	IF pSpan <> 0 THEN
		THIS^.AssertEquals_UDINT(2, pSpan^.links.count, 'Expected two links');
		THIS^.AssertTrue(pSpan^.parentSpanId = 0, 'Expected a link not to make the span a child');
		pSpan^.links.reset();
		pLink := pSpan^.links.next();
		THIS^.AssertTrue(
			pLink <> 0 AND_THEN pTrigger <> 0 AND_THEN MEMCMP(ADR(pLink^.spanId^.bytes), ADR(pTrigger^.spanId^.bytes), SIZEOF(spanId.bytes)) = 0,
			'Expected the first link to point at the trigger span'
		);
		pLink := pSpan^.links.next();
		THIS^.AssertTrue(pLink <> 0 AND_THEN pLink^.traceId^.bytes[0] = 16#AA, 'Expected the second link to point at the remote trace');
		pSpan^.delete(pSelf:=pSpan);
	END_IF
	IF pTrigger <> 0 THEN pTrigger^.delete(pSelf:=pTrigger); END_IF
TcUnit.TEST_FINISHED();
END_METHOD

(* A null or all zero link context fails the chain, and build then releases the span. *)
METHOD testRejectsInvalidLink : REFERENCE TO FB_Test
VAR
	resource: FB_Resource('');
	idGenerator: FB_MockIdGenerator;
	provider: FB_TracerProvider(resource:=resource, idGenerator:=idGenerator, sampler:=TcOtlp_GVL.defaultSampler);
	scope: FB_InstrumentationScope('tracer.test', '1.0.0', '');
	tracer: FB_Tracer(scope:=scope, provider:=provider);
	pSpan: POINTER TO FB_Span;
	pZero: POINTER TO FB_SpanContext;
	traceId: FB_TraceId;
	spanId: FB_SpanId;
	success: BOOL;
	reason: E_TracerFailureReason;
END_VAR
TcUnit.TEST('testRejectsInvalidLink');
	success := tracer.startSpan(name:='work').addLink(pContext:=0).build(pDest:=pSpan, failureReason=>reason);
	THIS^.AssertFalse(success, 'Expected a null link context to fail the chain');
	THIS^.AssertEquals_UDINT(TO_UDINT(E_TracerFailureReason.LINK_CONTEXT_POINTER_NULL), TO_UDINT(reason), 'Expected LINK_CONTEXT_POINTER_NULL');
	THIS^.AssertTrue(pSpan = 0, 'Expected no span');

	ContextFactory.buildContext(pDest:=pZero, pTraceId:=ADR(traceId), pSpanId:=ADR(spanId), pTraceState:=0, traceFlags:=0);
	success := tracer.startSpan(name:='work').addLink(pContext:=pZero).build(pDest:=pSpan, failureReason=>reason);
	THIS^.AssertFalse(success, 'Expected an all zero link context to fail the chain');
	THIS^.AssertEquals_UDINT(TO_UDINT(E_TracerFailureReason.LINK_CONTEXT_INVALID), TO_UDINT(reason), 'Expected LINK_CONTEXT_INVALID');
	THIS^.AssertTrue(pSpan = 0, 'Expected no span');

	IF pZero <> 0 THEN pZero^.delete(pSelf:=pZero); END_IF
	IF pSpan <> 0 THEN pSpan^.delete(pSelf:=pSpan); END_IF
TcUnit.TEST_FINISHED();
END_METHOD

END_FUNCTION_BLOCK

// ---- TEST/TRACING/PROCESSOR/FB_SpanProcessor_ForInspection.TcPOU
(* Processor test double that counts what the simple processor does with each span. *)
FUNCTION_BLOCK FB_SpanProcessor_ForInspection EXTENDS FB_SpanProcessor_Simple
VAR_OUTPUT
	enrichedCount: UDINT;
	exportedCount: UDINT;
	tickCount: UDINT;
	enrichedBeforeExport: BOOL;
	lastSpanName: T_MaxString;
END_VAR

METHOD enrich
VAR_IN_OUT
	span: FB_Span;
END_VAR
THIS^.enrichedCount := THIS^.enrichedCount + 1;
END_METHOD

METHOD export
VAR_INPUT
	span: REFERENCE TO FB_Span;
END_VAR
THIS^.exportedCount := THIS^.exportedCount + 1;
THIS^.enrichedBeforeExport := THIS^.enrichedCount = THIS^.exportedCount;
IF span.name <> 0 AND_THEN span.name^.pString <> 0 THEN
	THIS^.lastSpanName := span.name^.pString^;
END_IF
END_METHOD

METHOD tick
THIS^.tickCount := THIS^.tickCount + 1;
END_METHOD

END_FUNCTION_BLOCK

// ---- TEST/TRACING/SPAN/FB_TestSpanQueue.TcPOU
(* Tests FB_SpanQueue ordering, its bound, and the ownership hand-off on push and pop.

   The spans are opaque queue nodes: the queue only moves and releases pointers, so the tests
   allocate bare spans with __NEW instead of building them through FB_Tracer. *)
FUNCTION_BLOCK FB_TestSpanQueue EXTENDS FB_TestSuite

THIS^.testPushPopIsFifo();
THIS^.testPushDropsOldestWhenFull();
THIS^.testPopIntoAssignedDestinationFails();
THIS^.testCursorWalksWithoutTakingOwnership();
THIS^.testTransferToMovesOldestSpans();
THIS^.testTransferToRejectsInvalidDestination();
THIS^.testRotateMovesOldestToBack();

(* push takes ownership and clears the caller's pointer; pop returns spans oldest first. *)
METHOD testPushPopIsFifo : REFERENCE TO FB_Test
VAR
	queue: FB_SpanQueue(maxCount:=4);
	pFirst: POINTER TO FB_Span;
	pSecond: POINTER TO FB_Span;
	pExpectedFirst: POINTER TO FB_Span;
	pExpectedSecond: POINTER TO FB_Span;
	pPopped: POINTER TO FB_Span;
	reason: E_SpanQueueFailureReason;
END_VAR
TcUnit.TEST('testPushPopIsFifo');
	pFirst := __NEW(FB_Span);  // opaque queue node: the queue needs no span identity
	pSecond := __NEW(FB_Span);
	pExpectedFirst := pFirst;
	pExpectedSecond := pSecond;

	THIS^.AssertTrue(queue.push(pValue:=pFirst, failureReason=>reason), 'Expected the first push to succeed');
	THIS^.AssertTrue(queue.push(pValue:=pSecond, failureReason=>reason), 'Expected the second push to succeed');
	THIS^.AssertTrue(pFirst = 0 AND pSecond = 0, 'Expected push to clear the caller$'s pointers');
	THIS^.AssertEquals_UDINT(2, queue.count, 'Expected two queued spans');

	THIS^.AssertTrue(queue.pop(pValue:=pPopped, failureReason=>reason), 'Expected the first pop to succeed');
	THIS^.AssertTrue(pPopped = pExpectedFirst, 'Expected the oldest span first');
	IF pPopped <> 0 THEN pPopped^.delete(pSelf:=pPopped); END_IF

	THIS^.AssertTrue(queue.pop(pValue:=pPopped, failureReason=>reason), 'Expected the second pop to succeed');
	THIS^.AssertTrue(pPopped = pExpectedSecond, 'Expected the newer span second');
	IF pPopped <> 0 THEN pPopped^.delete(pSelf:=pPopped); END_IF

	THIS^.AssertFalse(queue.pop(pValue:=pPopped, failureReason=>reason), 'Expected pop on an empty queue to fail');
	THIS^.AssertEquals_UDINT(
		TO_UDINT(E_SpanQueueFailureReason.QUEUE_EMPTY),
		TO_UDINT(reason),
		'Expected QUEUE_EMPTY'
	);
	THIS^.AssertEquals_UDINT(0, queue.count, 'Expected the queue to be empty');
TcUnit.TEST_FINISHED();
END_METHOD

(* A full queue releases its oldest span to make room and counts the drop. *)
METHOD testPushDropsOldestWhenFull : REFERENCE TO FB_Test
VAR
	queue: FB_SpanQueue(maxCount:=1);
	pOld: POINTER TO FB_Span;
	pNew: POINTER TO FB_Span;
	pExpected: POINTER TO FB_Span;
	pPopped: POINTER TO FB_Span;
	reason: E_SpanQueueFailureReason;
END_VAR
TcUnit.TEST('testPushDropsOldestWhenFull');
	pOld := __NEW(FB_Span);  // opaque queue node: the queue needs no span identity
	pNew := __NEW(FB_Span);
	pExpected := pNew;

	queue.push(pValue:=pOld, failureReason=>reason);
	THIS^.AssertTrue(queue.push(pValue:=pNew, failureReason=>reason), 'Expected push to a full queue to succeed');
	THIS^.AssertEquals_UDINT(1, queue.count, 'Expected the bound to hold');
	THIS^.AssertEquals_UDINT(1, queue.droppedCount, 'Expected one dropped span');

	queue.pop(pValue:=pPopped, failureReason=>reason);
	THIS^.AssertTrue(pPopped = pExpected, 'Expected the newest span to be kept');
	IF pPopped <> 0 THEN pPopped^.delete(pSelf:=pPopped); END_IF
TcUnit.TEST_FINISHED();
END_METHOD

(* pop never overwrites a pointer the caller already owns, and free releases what is left. *)
METHOD testPopIntoAssignedDestinationFails : REFERENCE TO FB_Test
VAR
	queue: FB_SpanQueue(maxCount:=4);
	pQueued: POINTER TO FB_Span;
	pOwned: POINTER TO FB_Span;
	pExpected: POINTER TO FB_Span;
	reason: E_SpanQueueFailureReason;
END_VAR
TcUnit.TEST('testPopIntoAssignedDestinationFails');
	pQueued := __NEW(FB_Span);  // opaque queue node: the queue needs no span identity
	pOwned := __NEW(FB_Span);  // held by the caller, so pop must not overwrite it
	pExpected := pOwned;
	queue.push(pValue:=pQueued, failureReason=>reason);

	THIS^.AssertFalse(queue.pop(pValue:=pOwned, failureReason=>reason), 'Expected pop into an assigned pointer to fail');
	THIS^.AssertEquals_UDINT(
		TO_UDINT(E_SpanQueueFailureReason.DESTINATION_ALREADY_ASSIGNED),
		TO_UDINT(reason),
		'Expected DESTINATION_ALREADY_ASSIGNED'
	);
	THIS^.AssertTrue(pOwned = pExpected, 'Expected the destination to be left alone');
	THIS^.AssertEquals_UDINT(1, queue.count, 'Expected the span to stay queued');

	THIS^.AssertTrue(queue.free(), 'Expected free to release every span');
	THIS^.AssertEquals_UDINT(0, queue.count, 'Expected an empty queue after free');
	IF pOwned <> 0 THEN pOwned^.delete(pSelf:=pOwned); END_IF
TcUnit.TEST_FINISHED();
END_METHOD

(* reset and next walk the spans oldest first and leave them queued; pop keeps the cursor valid. *)
METHOD testCursorWalksWithoutTakingOwnership : REFERENCE TO FB_Test
VAR
	queue: FB_SpanQueue(maxCount:=4);
	pFirst: POINTER TO FB_Span;
	pSecond: POINTER TO FB_Span;
	pExpectedFirst: POINTER TO FB_Span;
	pExpectedSecond: POINTER TO FB_Span;
	pPopped: POINTER TO FB_Span;
END_VAR
TcUnit.TEST('testCursorWalksWithoutTakingOwnership');
	pFirst := __NEW(FB_Span);  // opaque queue node: the queue needs no span identity
	pSecond := __NEW(FB_Span);
	pExpectedFirst := pFirst;
	pExpectedSecond := pSecond;
	queue.push(pValue:=pFirst);
	queue.push(pValue:=pSecond);

	queue.reset();
	THIS^.AssertTrue(queue.next() = pExpectedFirst, 'Expected the oldest span first');
	THIS^.AssertTrue(queue.next() = pExpectedSecond, 'Expected the second span next');
	THIS^.AssertTrue(queue.next() = 0, 'Expected 0 after the last span');
	THIS^.AssertEquals_UDINT(2, queue.count, 'Expected the walk to leave both spans queued');

	// popping the node under the cursor moves the cursor to the new head
	queue.reset();
	queue.pop(pValue:=pPopped);
	THIS^.AssertTrue(queue.next() = pExpectedSecond, 'Expected the cursor to move past the popped span');

	IF pPopped <> 0 THEN pPopped^.delete(pSelf:=pPopped); END_IF
	queue.free();
	queue.reset();
	THIS^.AssertTrue(queue.next() = 0, 'Expected an empty walk after free');
TcUnit.TEST_FINISHED();
END_METHOD

(* transferTo moves the oldest spans, up to the destination's bound, without copying them. *)
METHOD testTransferToMovesOldestSpans : REFERENCE TO FB_Test
VAR
	source: FB_SpanQueue(maxCount:=4);
	destination: FB_SpanQueue(maxCount:=2);
	p: POINTER TO FB_Span;
	pFirst: POINTER TO FB_Span;
	pSecond: POINTER TO FB_Span;
	pThird: POINTER TO FB_Span;
	pPopped: POINTER TO FB_Span;
	reason: E_SpanQueueFailureReason;
END_VAR
TcUnit.TEST('testTransferToMovesOldestSpans');
	// opaque queue nodes: the queue needs no span identity
	p := __NEW(FB_Span); pFirst := p; source.push(pValue:=p, failureReason=>reason);
	p := __NEW(FB_Span); pSecond := p; source.push(pValue:=p, failureReason=>reason);
	p := __NEW(FB_Span); pThird := p; source.push(pValue:=p, failureReason=>reason);

	// ask for more than the destination's bound of 2 and more than the source holds
	THIS^.AssertTrue(source.transferTo(destination:=destination, count:=5, failureReason=>reason), 'Expected transferTo to succeed');
	THIS^.AssertEquals_UDINT(2, destination.count, 'Expected the destination bound to hold');
	THIS^.AssertEquals_UDINT(1, source.count, 'Expected one span left behind');

	destination.pop(pValue:=pPopped, failureReason=>reason);
	THIS^.AssertTrue(pPopped = pFirst, 'Expected the oldest span first');
	IF pPopped <> 0 THEN pPopped^.delete(pSelf:=pPopped); END_IF
	destination.pop(pValue:=pPopped, failureReason=>reason);
	THIS^.AssertTrue(pPopped = pSecond, 'Expected the second span next');
	IF pPopped <> 0 THEN pPopped^.delete(pSelf:=pPopped); END_IF
	source.pop(pValue:=pPopped, failureReason=>reason);
	THIS^.AssertTrue(pPopped = pThird, 'Expected the newest span to stay in the source');
	IF pPopped <> 0 THEN pPopped^.delete(pSelf:=pPopped); END_IF

	THIS^.AssertTrue(source.transferTo(destination:=destination, count:=1, failureReason=>reason), 'Expected an empty transfer to succeed');
	THIS^.AssertEquals_UDINT(0, destination.count, 'Expected nothing to move from an empty queue');
	source.free();
	destination.free();
TcUnit.TEST_FINISHED();
END_METHOD

(* transferTo refuses itself and a non-empty destination, and moves nothing. *)
METHOD testTransferToRejectsInvalidDestination : REFERENCE TO FB_Test
VAR
	source: FB_SpanQueue(maxCount:=4);
	destination: FB_SpanQueue(maxCount:=4);
	p: POINTER TO FB_Span;
	reason: E_SpanQueueFailureReason;
END_VAR
TcUnit.TEST('testTransferToRejectsInvalidDestination');
	// opaque queue nodes: the queue needs no span identity
	p := __NEW(FB_Span); source.push(pValue:=p, failureReason=>reason);
	p := __NEW(FB_Span); destination.push(pValue:=p, failureReason=>reason);  // makes the destination non-empty

	THIS^.AssertFalse(source.transferTo(destination:=source, count:=1, failureReason=>reason), 'Expected a self transfer to fail');
	THIS^.AssertEquals_UDINT(
		TO_UDINT(E_SpanQueueFailureReason.SELF_TRANSFER_NOT_ALLOWED),
		TO_UDINT(reason),
		'Expected SELF_TRANSFER_NOT_ALLOWED'
	);
	THIS^.AssertFalse(source.transferTo(destination:=destination, count:=1, failureReason=>reason), 'Expected a non-empty destination to fail');
	THIS^.AssertEquals_UDINT(
		TO_UDINT(E_SpanQueueFailureReason.DESTINATION_NOT_EMPTY),
		TO_UDINT(reason),
		'Expected DESTINATION_NOT_EMPTY'
	);
	THIS^.AssertTrue(source.count = 1 AND destination.count = 1, 'Expected both queues to be unchanged');
	source.free();
	destination.free();
TcUnit.TEST_FINISHED();
END_METHOD

(* rotate moves the oldest span to the back without releasing it, and fails on an empty queue. *)
METHOD testRotateMovesOldestToBack : REFERENCE TO FB_Test
VAR
	queue: FB_SpanQueue(maxCount:=0);  // 0 means the default bound, MAX_LOOP_COUNT
	pSpan: POINTER TO FB_Span;
	pFirst: POINTER TO FB_Span;
	pSecond: POINTER TO FB_Span;
	pPopped: POINTER TO FB_Span;
	reason: E_SpanQueueFailureReason;
END_VAR
TcUnit.TEST('testRotateMovesOldestToBack');
	THIS^.AssertFalse(queue.rotate(failureReason=>reason), 'Expected rotate on an empty queue to fail');
	THIS^.AssertEquals_UDINT(TO_UDINT(E_SpanQueueFailureReason.QUEUE_EMPTY), TO_UDINT(reason), 'Expected QUEUE_EMPTY');

	pSpan := __NEW(FB_Span);  // opaque queue node: the queue needs no span identity
	pFirst := pSpan;
	queue.push(pValue:=pSpan);
	pSpan := __NEW(FB_Span);
	pSecond := pSpan;
	queue.push(pValue:=pSpan);

	THIS^.AssertTrue(queue.rotate(failureReason=>reason), 'Expected rotate to succeed');
	THIS^.AssertEquals_UDINT(2, queue.count, 'Expected rotate to keep both spans');
	THIS^.AssertTrue(queue.next() = pSecond, 'Expected the cursor at the new head');
	queue.pop(pValue:=pPopped);
	THIS^.AssertTrue(pPopped = pSecond, 'Expected the second span first after a rotate');
	IF pPopped <> 0 THEN pPopped^.delete(pSelf:=pPopped); END_IF
	queue.pop(pValue:=pPopped);
	THIS^.AssertTrue(pPopped = pFirst, 'Expected the rotated span last');
	IF pPopped <> 0 THEN pPopped^.delete(pSelf:=pPopped); END_IF
	queue.free();
TcUnit.TEST_FINISHED();
END_METHOD

END_FUNCTION_BLOCK

// ---- TEST/TRACING/PROCESSOR/FB_TestSpanProcessors.TcPOU
(* Tests FB_SpanProcessor_Simple and FB_SpanProcessor_Batch and their hand-off to an exporter. *)
FUNCTION_BLOCK FB_TestSpanProcessors EXTENDS FB_TestSuite
VAR
	// kept across scans by testBatchExportsAfterScheduledDelay
	_resource: FB_Resource('');
	_idGenerator: FB_MockIdGenerator;
	_provider: FB_TracerProvider_ForInspection(resource:=_resource, idGenerator:=_idGenerator, sampler:=TcOtlp_GVL.defaultSampler);
	_scope: FB_InstrumentationScope('tracer.test', '1.0.0', '');
	_tracer: FB_Tracer(scope:=_scope, provider:=_provider);
	_exporter: FB_SpanExporter_ForInspection;
	_processor: FB_SpanProcessor_Batch(maxQueueSize:=10, scheduledDelayMillis:=50, maxExportBatchSize:=10, exporter:=_exporter);
END_VAR

THIS^.testSimpleEnrichesThenExports();
THIS^.testSimpleHandsCloneToExporter();
THIS^.testSimpleDropsSpanWhenExporterBusy();
THIS^.testBatchWaitsForFullBatch();
THIS^.testBatchKeepsSpansWhileExporterBusy();
THIS^.testBatchDropsOldestWhenFull();
THIS^.testBatchIgnoresSpansWithoutExporter();
THIS^.testBatchExportsAfterScheduledDelay();

(* The simple processor enriches each span and then exports it, once per span. *)
METHOD testSimpleEnrichesThenExports : REFERENCE TO FB_Test
VAR
	resource: FB_Resource('');
	idGenerator: FB_MockIdGenerator;
	provider: FB_TracerProvider_ForInspection(resource:=resource, idGenerator:=idGenerator, sampler:=TcOtlp_GVL.defaultSampler);
	scope: FB_InstrumentationScope('tracer.test', '1.0.0', '');
	tracer: FB_Tracer(scope:=scope, provider:=provider);
	processor: FB_SpanProcessor_ForInspection(exporter:=0);
	pSpan: POINTER TO FB_Span;
END_VAR
TcUnit.TEST('testSimpleEnrichesThenExports');
	tracer.startSpan(name:='work').build(pDest:=pSpan);
	THIS^.AssertTrue(pSpan <> 0, 'Expected the span to build');
	IF pSpan <> 0 THEN
		processor.onEnd(pSpan^);
		pSpan^.delete(pSelf:=pSpan);
	END_IF
	THIS^.AssertEquals_UDINT(1, processor.enrichedCount, 'Expected one enrich');
	THIS^.AssertEquals_UDINT(1, processor.exportedCount, 'Expected one export');
	THIS^.AssertTrue(processor.enrichedBeforeExport, 'Expected enrich to run before export');
	THIS^.AssertEquals_STRING('work', processor.lastSpanName, 'Expected the span to be exported');
TcUnit.TEST_FINISHED();
END_METHOD

(* The simple processor gives the exporter a clone, which outlives the span the provider releases. *)
METHOD testSimpleHandsCloneToExporter : REFERENCE TO FB_Test
VAR
	resource: FB_Resource('');
	idGenerator: FB_MockIdGenerator;
	provider: FB_TracerProvider_ForInspection(resource:=resource, idGenerator:=idGenerator, sampler:=TcOtlp_GVL.defaultSampler);
	scope: FB_InstrumentationScope('tracer.test', '1.0.0', '');
	tracer: FB_Tracer(scope:=scope, provider:=provider);
	exporter: FB_SpanExporter_ForInspection;
	processor: FB_SpanProcessor_Simple(exporter:=exporter);
	pSpan: POINTER TO FB_Span;
	pSource: POINTER TO FB_Span;
	pHeld: POINTER TO FB_Span;
END_VAR
TcUnit.TEST('testSimpleHandsCloneToExporter');
	tracer.startSpan(name:='work').build(pDest:=pSpan);
	THIS^.AssertTrue(pSpan <> 0, 'Expected the span to build');
	IF pSpan <> 0 THEN
		pSource := pSpan;
		processor.onEnd(pSpan^);
		pSpan^.delete(pSelf:=pSpan);
	END_IF
	THIS^.AssertEquals_UDINT(1, exporter.exportCount, 'Expected one export');
	THIS^.AssertEquals_UDINT(1, exporter.lastBatchCount, 'Expected a batch of one');
	pHeld := exporter.heldSpan();
	THIS^.AssertTrue(pHeld <> 0 AND_THEN pHeld <> pSource, 'Expected the exporter to hold a clone');
	IF pHeld <> 0 AND_THEN pHeld^.name <> 0 THEN
		THIS^.AssertEquals_STRING('work', pHeld^.name^.pString^, 'Expected the clone to outlive the source');
	END_IF
	processor.tick();
	THIS^.AssertEquals_UDINT(1, exporter.tickCount, 'Expected tick to reach the exporter');
	exporter.free();
TcUnit.TEST_FINISHED();
END_METHOD

(* A busy exporter is not offered the span, and nothing is kept for later. *)
METHOD testSimpleDropsSpanWhenExporterBusy : REFERENCE TO FB_Test
VAR
	resource: FB_Resource('');
	idGenerator: FB_MockIdGenerator;
	provider: FB_TracerProvider_ForInspection(resource:=resource, idGenerator:=idGenerator, sampler:=TcOtlp_GVL.defaultSampler);
	scope: FB_InstrumentationScope('tracer.test', '1.0.0', '');
	tracer: FB_Tracer(scope:=scope, provider:=provider);
	exporter: FB_SpanExporter_ForInspection;
	processor: FB_SpanProcessor_Simple(exporter:=exporter);
	pSpan: POINTER TO FB_Span;
END_VAR
TcUnit.TEST('testSimpleDropsSpanWhenExporterBusy');
	exporter.busy := TRUE;
	tracer.startSpan(name:='work').build(pDest:=pSpan);
	IF pSpan <> 0 THEN
		processor.onEnd(pSpan^);
		pSpan^.delete(pSelf:=pSpan);
	END_IF
	THIS^.AssertEquals_UDINT(0, exporter.exportCount, 'Expected no export while busy');
	THIS^.AssertEquals_UDINT(0, exporter.callsWhileBusy, 'Expected the processor not to call a busy exporter');
	THIS^.AssertTrue(exporter.heldSpan() = 0, 'Expected the exporter to hold nothing');
TcUnit.TEST_FINISHED();
END_METHOD

(* Ended spans are only queued; a full batch goes out on the next tick without waiting for the delay. *)
METHOD testBatchWaitsForFullBatch : REFERENCE TO FB_Test
VAR
	resource: FB_Resource('');
	idGenerator: FB_MockIdGenerator;
	provider: FB_TracerProvider_ForInspection(resource:=resource, idGenerator:=idGenerator, sampler:=TcOtlp_GVL.defaultSampler);
	scope: FB_InstrumentationScope('tracer.test', '1.0.0', '');
	tracer: FB_Tracer(scope:=scope, provider:=provider);
	exporter: FB_SpanExporter_ForInspection;
	processor: FB_SpanProcessor_Batch(maxQueueSize:=10, scheduledDelayMillis:=60000, maxExportBatchSize:=3, exporter:=exporter);
	pSpan: POINTER TO FB_Span;
END_VAR
TcUnit.TEST('testBatchWaitsForFullBatch');
	tracer.startSpan(name:='a').build(pDest:=pSpan);
	IF pSpan <> 0 THEN
		processor.onEnd(pSpan^);
		pSpan^.delete(pSelf:=pSpan);
	END_IF
	tracer.startSpan(name:='b').build(pDest:=pSpan);
	IF pSpan <> 0 THEN
		processor.onEnd(pSpan^);
		pSpan^.delete(pSelf:=pSpan);
	END_IF
	THIS^.AssertEquals_UDINT(0, exporter.exportCount, 'Expected onEnd not to export');
	THIS^.AssertEquals_UDINT(2, processor.queuedCount, 'Expected two queued spans');
	processor.tick();
	THIS^.AssertEquals_UDINT(0, exporter.exportCount, 'Expected no export before a full batch or the delay');
	THIS^.AssertEquals_UDINT(1, exporter.tickCount, 'Expected tick to reach the exporter');
	tracer.startSpan(name:='c').build(pDest:=pSpan);
	IF pSpan <> 0 THEN
		processor.onEnd(pSpan^);
		pSpan^.delete(pSelf:=pSpan);
	END_IF
	processor.tick();
	THIS^.AssertEquals_UDINT(1, exporter.exportCount, 'Expected one export for the full batch');
	THIS^.AssertEquals_UDINT(3, exporter.lastBatchCount, 'Expected the three spans in one batch');
	THIS^.AssertEquals_UDINT(0, processor.queuedCount, 'Expected the queue to be empty');
	THIS^.AssertEquals_UDINT(0, processor.droppedCount, 'Expected nothing dropped');
	exporter.free();
	processor.free();
TcUnit.TEST_FINISHED();
END_METHOD

(* Spans that end while the exporter is busy stay queued and are exported once it is idle. *)
METHOD testBatchKeepsSpansWhileExporterBusy : REFERENCE TO FB_Test
VAR
	resource: FB_Resource('');
	idGenerator: FB_MockIdGenerator;
	provider: FB_TracerProvider_ForInspection(resource:=resource, idGenerator:=idGenerator, sampler:=TcOtlp_GVL.defaultSampler);
	scope: FB_InstrumentationScope('tracer.test', '1.0.0', '');
	tracer: FB_Tracer(scope:=scope, provider:=provider);
	exporter: FB_SpanExporter_ForInspection;
	processor: FB_SpanProcessor_Batch(maxQueueSize:=10, scheduledDelayMillis:=60000, maxExportBatchSize:=1, exporter:=exporter);
	pSpan: POINTER TO FB_Span;
	pHeld: POINTER TO FB_Span;
END_VAR
TcUnit.TEST('testBatchKeepsSpansWhileExporterBusy');
	exporter.busy := TRUE;
	tracer.startSpan(name:='first').build(pDest:=pSpan);
	IF pSpan <> 0 THEN
		processor.onEnd(pSpan^);
		pSpan^.delete(pSelf:=pSpan);
	END_IF
	tracer.startSpan(name:='second').build(pDest:=pSpan);
	IF pSpan <> 0 THEN
		processor.onEnd(pSpan^);
		pSpan^.delete(pSelf:=pSpan);
	END_IF
	processor.tick();
	THIS^.AssertEquals_UDINT(0, exporter.exportCount, 'Expected no export while busy');
	THIS^.AssertEquals_UDINT(0, exporter.callsWhileBusy, 'Expected the processor not to call a busy exporter');
	THIS^.AssertEquals_UDINT(2, processor.queuedCount, 'Expected both spans kept');

	exporter.busy := FALSE;
	processor.tick();
	THIS^.AssertEquals_UDINT(1, exporter.exportCount, 'Expected an export once idle');
	THIS^.AssertEquals_UDINT(1, exporter.lastBatchCount, 'Expected a batch of maxExportBatchSize');
	pHeld := exporter.heldSpan();
	IF pHeld <> 0 AND_THEN pHeld^.name <> 0 THEN
		THIS^.AssertEquals_STRING('first', pHeld^.name^.pString^, 'Expected the oldest span first');
	ELSE
		THIS^.AssertTrue(FALSE, 'Expected the exporter to hold a span');
	END_IF
	THIS^.AssertEquals_UDINT(1, processor.queuedCount, 'Expected the newer span to wait');

	processor.tick();
	THIS^.AssertEquals_UDINT(2, exporter.exportCount, 'Expected the second span on the next tick');
	pHeld := exporter.heldSpan();
	IF pHeld <> 0 AND_THEN pHeld^.name <> 0 THEN
		THIS^.AssertEquals_STRING('second', pHeld^.name^.pString^, 'Expected the newer span second');
	END_IF
	THIS^.AssertEquals_UDINT(0, processor.droppedCount, 'Expected nothing dropped');
	exporter.free();
	processor.free();
TcUnit.TEST_FINISHED();
END_METHOD

(* A full queue drops its oldest span for the newest and counts it. *)
METHOD testBatchDropsOldestWhenFull : REFERENCE TO FB_Test
VAR
	resource: FB_Resource('');
	idGenerator: FB_MockIdGenerator;
	provider: FB_TracerProvider_ForInspection(resource:=resource, idGenerator:=idGenerator, sampler:=TcOtlp_GVL.defaultSampler);
	scope: FB_InstrumentationScope('tracer.test', '1.0.0', '');
	tracer: FB_Tracer(scope:=scope, provider:=provider);
	exporter: FB_SpanExporter_ForInspection;
	processor: FB_SpanProcessor_Batch(maxQueueSize:=2, scheduledDelayMillis:=60000, maxExportBatchSize:=2, exporter:=exporter);
	pSpan: POINTER TO FB_Span;
	pHeld: POINTER TO FB_Span;
END_VAR
TcUnit.TEST('testBatchDropsOldestWhenFull');
	exporter.busy := TRUE;
	tracer.startSpan(name:='a').build(pDest:=pSpan);
	IF pSpan <> 0 THEN
		processor.onEnd(pSpan^);
		pSpan^.delete(pSelf:=pSpan);
	END_IF
	tracer.startSpan(name:='b').build(pDest:=pSpan);
	IF pSpan <> 0 THEN
		processor.onEnd(pSpan^);
		pSpan^.delete(pSelf:=pSpan);
	END_IF
	tracer.startSpan(name:='c').build(pDest:=pSpan);
	IF pSpan <> 0 THEN
		processor.onEnd(pSpan^);
		pSpan^.delete(pSelf:=pSpan);
	END_IF
	THIS^.AssertEquals_UDINT(2, processor.queuedCount, 'Expected the queue to stay at maxQueueSize');
	THIS^.AssertEquals_UDINT(1, processor.droppedCount, 'Expected one dropped span');
	processor.tick();
	THIS^.AssertEquals_UDINT(0, exporter.callsWhileBusy, 'Expected the processor not to call a busy exporter with a full batch');
	exporter.busy := FALSE;
	processor.tick();
	THIS^.AssertEquals_UDINT(2, exporter.lastBatchCount, 'Expected the two kept spans');
	pHeld := exporter.heldSpan();
	IF pHeld <> 0 AND_THEN pHeld^.name <> 0 THEN
		THIS^.AssertEquals_STRING('b', pHeld^.name^.pString^, 'Expected the oldest span to be the one dropped');
	ELSE
		THIS^.AssertTrue(FALSE, 'Expected the exporter to hold a span');
	END_IF
	exporter.free();
	processor.free();
TcUnit.TEST_FINISHED();
END_METHOD

(* With no exporter the processor keeps nothing. *)
METHOD testBatchIgnoresSpansWithoutExporter : REFERENCE TO FB_Test
VAR
	resource: FB_Resource('');
	idGenerator: FB_MockIdGenerator;
	provider: FB_TracerProvider_ForInspection(resource:=resource, idGenerator:=idGenerator, sampler:=TcOtlp_GVL.defaultSampler);
	scope: FB_InstrumentationScope('tracer.test', '1.0.0', '');
	tracer: FB_Tracer(scope:=scope, provider:=provider);
	exporter: FB_SpanExporter_ForInspection;
	processor: FB_SpanProcessor_Batch(maxQueueSize:=10, scheduledDelayMillis:=0, maxExportBatchSize:=1, exporter:=0);
	pSpan: POINTER TO FB_Span;
END_VAR
TcUnit.TEST('testBatchIgnoresSpansWithoutExporter');
	tracer.startSpan(name:='work').build(pDest:=pSpan);
	IF pSpan <> 0 THEN
		processor.onEnd(pSpan^);
		pSpan^.delete(pSelf:=pSpan);
	END_IF
	processor.tick();
	THIS^.AssertEquals_UDINT(0, processor.queuedCount, 'Expected nothing queued');
TcUnit.TEST_FINISHED();
END_METHOD

(* A partial batch is exported once scheduledDelayMillis has passed, and not before. *)
METHOD testBatchExportsAfterScheduledDelay : REFERENCE TO FB_Test
VAR CONSTANT
	DELAY_MILLIS: UDINT := 50;  // matches _processor's scheduledDelayMillis
	MAX_CYCLES: UDINT := 1000;
END_VAR
VAR_INST
	_started: BOOL;
	_finished: BOOL;
	_cycles: UDINT;
	_startTime: ULINT;
END_VAR
VAR
	pSpan: POINTER TO FB_Span;
	elapsedMillis: ULINT;
END_VAR
TcUnit.TEST('testBatchExportsAfterScheduledDelay');
	IF _finished THEN
		RETURN;
	END_IF
	IF NOT _started THEN
		_tracer.startSpan(name:='work').build(pDest:=pSpan);
		IF pSpan <> 0 THEN
			_processor.onEnd(pSpan^);
			pSpan^.delete(pSelf:=pSpan);
		END_IF
		_startTime := F_GetSystemTime();
		_started := TRUE;
	END_IF

	_processor.tick();
	_cycles := _cycles + 1;
	IF _exporter.exportCount > 0 OR _cycles > MAX_CYCLES THEN
		elapsedMillis := (F_GetSystemTime() - _startTime) / 10000;  // 100 ns ticks
		THIS^.AssertEquals_UDINT(1, _exporter.exportCount, 'Expected the partial batch to be exported');
		THIS^.AssertEquals_UDINT(1, _exporter.lastBatchCount, 'Expected a batch of one');
		THIS^.AssertTrue(elapsedMillis >= DELAY_MILLIS - 1, 'Expected the export to wait for the delay');
		_exporter.free();
		_processor.free();
		_finished := TRUE;
		TcUnit.TEST_FINISHED();
	END_IF
END_METHOD

END_FUNCTION_BLOCK

// ---- TEST/TRACING/EXPORTING/FB_SpanExporter_ForInspection.TcPOU
(*
	Span exporter test double. It keeps each accepted batch until the next one or free, and is
	busy while busy is set. callsWhileBusy counts export calls made while busy, which a processor
	must never make.
*)
FUNCTION_BLOCK FB_SpanExporter_ForInspection EXTENDS FB_SpanExporter_Base
VAR_INPUT
	busy: BOOL;
END_VAR
VAR_OUTPUT
	exportCount: UDINT;
	lastBatchCount: UDINT;
	tickCount: UDINT;
	callsWhileBusy: UDINT;
END_VAR

METHOD export : BOOL
VAR_IN_OUT
	spans: FB_SpanQueue;
END_VAR
VAR_INPUT
	count: UDINT;
END_VAR
VAR_OUTPUT
	failureReason: E_SpanExporterFailureReason;
END_VAR
IF THIS^.isBusy() THEN
	THIS^.callsWhileBusy := THIS^.callsWhileBusy + 1;
END_IF
export := SUPER^.export(spans:=spans, count:=count, failureReason=>failureReason);
IF export THEN
	THIS^.exportCount := THIS^.exportCount + 1;
	THIS^.lastBatchCount := THIS^._spans.count;
	// nothing is delivered, so the batch stays held until the next one or free
	THIS^._exportActive := FALSE;
END_IF
END_METHOD

(* The oldest span of the held batch, borrowed; 0 when nothing is held. *)
METHOD heldSpan : POINTER TO FB_Span
THIS^._spans.reset();
heldSpan := THIS^._spans.next();
END_METHOD

METHOD isBusy : BOOL
isBusy := THIS^.busy;
END_METHOD

METHOD tick : BOOL
VAR_OUTPUT
	failureReason: E_SpanExporterFailureReason;
END_VAR
THIS^.tickCount := THIS^.tickCount + 1;
failureReason := E_SpanExporterFailureReason.NA;
tick := TRUE;
END_METHOD

END_FUNCTION_BLOCK

// ---- TEST/TRACING/PROVIDER/FB_TestTracerProvider.TcPOU
(* Tests FB_TracerProvider processor staging and the hand-over of ended spans in tick. *)
FUNCTION_BLOCK FB_TestTracerProvider EXTENDS FB_TestSuite

THIS^.testTickHandsSpansToEachProcessor();
THIS^.testStageProcessorIgnoresDuplicates();
THIS^.testTickWithoutProcessorsSucceeds();
THIS^.testProcessorsMustBeStagedEachScan();

(* Every staged processor receives every ended span once; tick then releases the spans. *)
METHOD testTickHandsSpansToEachProcessor : REFERENCE TO FB_Test
VAR
	resource: FB_Resource('');
	idGenerator: FB_MockIdGenerator;
	provider: FB_TracerProvider_ForInspection(resource:=resource, idGenerator:=idGenerator, sampler:=TcOtlp_GVL.defaultSampler);
	scope: FB_InstrumentationScope('tracer.test', '1.0.0', '');
	tracer: FB_Tracer(scope:=scope, provider:=provider);
	processorA: FB_SpanProcessor_ForInspection(exporter:=0);
	processorB: FB_SpanProcessor_ForInspection(exporter:=0);
	pSpan: POINTER TO FB_Span;
	success: BOOL;
	reason: E_TracerProviderFailureReason;
END_VAR
TcUnit.TEST('testTickHandsSpansToEachProcessor');
	provider.stageProcessor(processorA).stageProcessor(processorB);
	tracer.startSpan(name:='first').build(pDest:=pSpan);
	tracer.endSpan(pSpan:=pSpan);
	tracer.startSpan(name:='second').build(pDest:=pSpan);
	tracer.endSpan(pSpan:=pSpan);

	success := provider.tick(failureReason=>reason);
	THIS^.AssertTrue(success, 'Expected tick to succeed');
	THIS^.AssertEquals_UDINT(
		TO_UDINT(E_TracerProviderFailureReason.NA),
		TO_UDINT(reason),
		'Expected no failure reason on success'
	);
	THIS^.AssertEquals_UDINT(2, processorA.exportedCount, 'Expected processor A to get both spans');
	THIS^.AssertEquals_UDINT(2, processorB.exportedCount, 'Expected processor B to get both spans');
	THIS^.AssertEquals_STRING('second', processorA.lastSpanName, 'Expected the spans in the order they ended');
	THIS^.AssertEquals_UDINT(1, processorA.tickCount, 'Expected each processor to be ticked once');
	THIS^.AssertEquals_UDINT(0, provider.spans.count, 'Expected the queue to be empty');
	THIS^.AssertEquals_UDINT(0, provider.stagedProcessorCount, 'Expected the staged list to be cleared');
TcUnit.TEST_FINISHED();
END_METHOD

(* Staging the same processor twice gives it each span once. *)
METHOD testStageProcessorIgnoresDuplicates : REFERENCE TO FB_Test
VAR
	resource: FB_Resource('');
	idGenerator: FB_MockIdGenerator;
	provider: FB_TracerProvider_ForInspection(resource:=resource, idGenerator:=idGenerator, sampler:=TcOtlp_GVL.defaultSampler);
	scope: FB_InstrumentationScope('tracer.test', '1.0.0', '');
	tracer: FB_Tracer(scope:=scope, provider:=provider);
	processor: FB_SpanProcessor_ForInspection(exporter:=0);
	pSpan: POINTER TO FB_Span;
END_VAR
TcUnit.TEST('testStageProcessorIgnoresDuplicates');
	provider.stageProcessor(processor).stageProcessor(processor);
	THIS^.AssertEquals_UDINT(1, provider.stagedProcessorCount, 'Expected the duplicate to be ignored');

	tracer.startSpan(name:='work').build(pDest:=pSpan);
	tracer.endSpan(pSpan:=pSpan);
	provider.tick();
	THIS^.AssertEquals_UDINT(1, processor.exportedCount, 'Expected the span exactly once');
TcUnit.TEST_FINISHED();
END_METHOD

(* With no processors staged, tick releases the queued spans and still succeeds. *)
METHOD testTickWithoutProcessorsSucceeds : REFERENCE TO FB_Test
VAR
	resource: FB_Resource('');
	idGenerator: FB_MockIdGenerator;
	provider: FB_TracerProvider_ForInspection(resource:=resource, idGenerator:=idGenerator, sampler:=TcOtlp_GVL.defaultSampler);
	scope: FB_InstrumentationScope('tracer.test', '1.0.0', '');
	tracer: FB_Tracer(scope:=scope, provider:=provider);
	pSpan: POINTER TO FB_Span;
	success: BOOL;
END_VAR
TcUnit.TEST('testTickWithoutProcessorsSucceeds');
	tracer.startSpan(name:='work').build(pDest:=pSpan);
	tracer.endSpan(pSpan:=pSpan);
	THIS^.AssertEquals_UDINT(1, provider.spans.count, 'Expected the span to be queued');

	success := provider.tick();
	THIS^.AssertTrue(success, 'Expected tick to succeed');
	THIS^.AssertEquals_UDINT(0, provider.spans.count, 'Expected tick to release the span');
TcUnit.TEST_FINISHED();
END_METHOD

(* tick clears the staged list, so a processor that is not staged again gets nothing. *)
METHOD testProcessorsMustBeStagedEachScan : REFERENCE TO FB_Test
VAR
	resource: FB_Resource('');
	idGenerator: FB_MockIdGenerator;
	provider: FB_TracerProvider_ForInspection(resource:=resource, idGenerator:=idGenerator, sampler:=TcOtlp_GVL.defaultSampler);
	scope: FB_InstrumentationScope('tracer.test', '1.0.0', '');
	tracer: FB_Tracer(scope:=scope, provider:=provider);
	processor: FB_SpanProcessor_ForInspection(exporter:=0);
	pSpan: POINTER TO FB_Span;
END_VAR
TcUnit.TEST('testProcessorsMustBeStagedEachScan');
	provider.stageProcessor(processor);
	provider.tick();

	tracer.startSpan(name:='work').build(pDest:=pSpan);
	tracer.endSpan(pSpan:=pSpan);
	provider.tick();
	THIS^.AssertEquals_UDINT(0, processor.exportedCount, 'Expected an unstaged processor to get nothing');
TcUnit.TEST_FINISHED();
END_METHOD

END_FUNCTION_BLOCK

// ---- TEST/TRACING/SAMPLING/FB_TestSamplers.TcPOU
(* Tests the span samplers: onStart makes the head decision when a span is built, and
   FB_TracerProvider asks onEnd only about spans that are still sampled. *)
FUNCTION_BLOCK FB_TestSamplers EXTENDS FB_TestSuite

THIS^.testDefaultSamplerFollowsParent();
THIS^.testAlwaysOnSamplesChildOfUnsampledParent();
THIS^.testErrorsOnlyKeepsFailedSpans();
THIS^.testOnEndCannotKeepSpanDroppedOnStart();
THIS^.testLinkDoesNotAffectSampling();

(* Builds a root span, or a child of pParent, gives it a status, and ends it. Returns endSpan's
   result, or FALSE when the span could not be built. *)
METHOD _endSpan : BOOL
VAR_INPUT
	tracer: REFERENCE TO FB_Tracer;
	name: T_MaxString;
	statusCode: E_StatusCode;
	pParent: POINTER TO FB_SpanContext;  // 0 for a root span
END_VAR
VAR
	_pSpan: POINTER TO FB_Span;
	_built: BOOL;
END_VAR
IF pParent = 0 THEN
	_built := tracer.startSpan(name:=name).build(pDest:=_pSpan);
ELSE
	_built := tracer.startSpan(name:=name).setParentUsingContext(pContext:=pParent).build(pDest:=_pSpan);
END_IF
IF NOT _built THEN
	RETURN;
END_IF

CASE statusCode OF
	E_StatusCode.STATUS_CODE_OK:
		tracer.setSpanStatusOk(pSpan:=_pSpan);
	E_StatusCode.STATUS_CODE_ERROR:
		tracer.setSpanStatusError(pSpan:=_pSpan, message:='boom');
END_CASE
_endSpan := tracer.endSpan(pSpan:=_pSpan);
END_METHOD

(* The default sampler is ParentBased(root=AlwaysOn): a root span is sampled, the child of a
   sampled remote parent is sampled, and the child of an unsampled one is not. Status does not
   matter to it. *)
METHOD testDefaultSamplerFollowsParent : REFERENCE TO FB_Test
VAR
	resource: FB_Resource('');
	idGenerator: FB_MockIdGenerator;
	provider: FB_TracerProvider_ForInspection(resource:=resource, idGenerator:=idGenerator, sampler:=TcOtlp_GVL.defaultSampler);
	scope: FB_InstrumentationScope('sampler.test', '1.0.0', '');
	tracer: FB_Tracer(scope:=scope, provider:=provider);
	processor: FB_SpanProcessor_ForInspection(exporter:=0);
	sampled: STRING(55) := '00-4bf92f3577b34da6a3ce929d0e0e4736-00f067aa0ba902b7-01';
	unsampled: STRING(55) := '00-4bf92f3577b34da6a3ce929d0e0e4736-00f067aa0ba902b7-00';
	pSampledParent: POINTER TO FB_SpanContext;
	pUnsampledParent: POINTER TO FB_SpanContext;
END_VAR
TcUnit.TEST('testDefaultSamplerFollowsParent');
	TraceContextPropagator.extract(pDest:=pSampledParent, traceparent:=sampled, tracestate:='');
	TraceContextPropagator.extract(pDest:=pUnsampledParent, traceparent:=unsampled, tracestate:='');
	THIS^.AssertTrue(pSampledParent <> 0 AND pUnsampledParent <> 0, 'Expected both parents to be extracted');

	provider.stageProcessor(processor);
	THIS^._endSpan(tracer:=tracer, name:='root.failed', statusCode:=E_StatusCode.STATUS_CODE_ERROR, pParent:=0);
	THIS^._endSpan(tracer:=tracer, name:='root.ok', statusCode:=E_StatusCode.STATUS_CODE_OK, pParent:=0);
	THIS^._endSpan(tracer:=tracer, name:='unsampled.child', statusCode:=E_StatusCode.STATUS_CODE_UNSET, pParent:=pUnsampledParent);
	THIS^._endSpan(tracer:=tracer, name:='sampled.child', statusCode:=E_StatusCode.STATUS_CODE_UNSET, pParent:=pSampledParent);
	provider.tick();

	THIS^.AssertEquals_UDINT(3, processor.exportedCount, 'Expected both roots and the sampled child to be processed');
	THIS^.AssertEquals_STRING('sampled.child', processor.lastSpanName, 'Expected the sampled child to be processed last');

	IF pSampledParent <> 0 THEN pSampledParent^.delete(pSelf:=pSampledParent); END_IF
	IF pUnsampledParent <> 0 THEN pUnsampledParent^.delete(pSelf:=pUnsampledParent); END_IF
TcUnit.TEST_FINISHED();
END_METHOD

(* The always-on sampler samples every span, even the child of a parent that was not sampled,
   and the decision is carried into the span's context. *)
METHOD testAlwaysOnSamplesChildOfUnsampledParent : REFERENCE TO FB_Test
VAR
	alwaysOn: FB_Sampler_AlwaysOn;
	resource: FB_Resource('');
	idGenerator: FB_MockIdGenerator;
	provider: FB_TracerProvider_ForInspection(resource:=resource, idGenerator:=idGenerator, sampler:=alwaysOn);
	scope: FB_InstrumentationScope('sampler.test', '1.0.0', '');
	tracer: FB_Tracer(scope:=scope, provider:=provider);
	processor: FB_SpanProcessor_ForInspection(exporter:=0);
	unsampled: STRING(55) := '00-4bf92f3577b34da6a3ce929d0e0e4736-00f067aa0ba902b7-00';
	pParent: POINTER TO FB_SpanContext;
	pSpan: POINTER TO FB_Span;
	pContext: POINTER TO FB_SpanContext;
END_VAR
TcUnit.TEST('testAlwaysOnSamplesChildOfUnsampledParent');
	TraceContextPropagator.extract(pDest:=pParent, traceparent:=unsampled, tracestate:='');
	THIS^.AssertTrue(pParent <> 0, 'Expected the unsampled parent to be extracted');

	provider.stageProcessor(processor);
	tracer.startSpan(name:='child').setParentUsingContext(pContext:=pParent).build(pDest:=pSpan);
	THIS^.AssertTrue(pSpan <> 0, 'Expected the child to be built');
	IF pSpan <> 0 THEN
		tracer.getSpanContext(pSpan:=pSpan, pDest:=pContext);
		THIS^.AssertTrue(pContext <> 0 AND_THEN (pContext^.traceFlags AND 16#01) <> 0, 'Expected the child$'s context to carry the sampled bit');
	END_IF
	tracer.endSpan(pSpan:=pSpan);
	provider.tick();

	THIS^.AssertEquals_UDINT(1, processor.exportedCount, 'Expected the child to be processed');

	IF pContext <> 0 THEN pContext^.delete(pSelf:=pContext); END_IF
	IF pParent <> 0 THEN pParent^.delete(pSelf:=pParent); END_IF
TcUnit.TEST_FINISHED();
END_METHOD

(* The errors-only sampler keeps a span that ended with an error status and releases the
   others. Dropping a span is not a failure, so endSpan still succeeds. *)
METHOD testErrorsOnlyKeepsFailedSpans : REFERENCE TO FB_Test
VAR
	errorsOnly: FB_Sampler_ErrorsOnly;
	resource: FB_Resource('');
	idGenerator: FB_MockIdGenerator;
	provider: FB_TracerProvider_ForInspection(resource:=resource, idGenerator:=idGenerator, sampler:=errorsOnly);
	scope: FB_InstrumentationScope('sampler.test', '1.0.0', '');
	tracer: FB_Tracer(scope:=scope, provider:=provider);
	processor: FB_SpanProcessor_ForInspection(exporter:=0);
	endedUnset: BOOL;
	endedOk: BOOL;
	endedFailed: BOOL;
END_VAR
TcUnit.TEST('testErrorsOnlyKeepsFailedSpans');
	provider.stageProcessor(processor);
	endedUnset := THIS^._endSpan(tracer:=tracer, name:='unset', statusCode:=E_StatusCode.STATUS_CODE_UNSET, pParent:=0);
	endedOk := THIS^._endSpan(tracer:=tracer, name:='ok', statusCode:=E_StatusCode.STATUS_CODE_OK, pParent:=0);
	endedFailed := THIS^._endSpan(tracer:=tracer, name:='failed', statusCode:=E_StatusCode.STATUS_CODE_ERROR, pParent:=0);

	THIS^.AssertTrue(endedUnset AND endedOk AND endedFailed, 'Expected endSpan to succeed for kept and dropped spans');
	THIS^.AssertEquals_UDINT(1, provider.spans.count, 'Expected only the failed span to be queued');

	provider.tick();
	THIS^.AssertEquals_UDINT(1, processor.exportedCount, 'Expected one span to reach the processor');
	THIS^.AssertEquals_STRING('failed', processor.lastSpanName, 'Expected the failed span to be the one kept');
TcUnit.TEST_FINISHED();
END_METHOD

(* A span dropped by onStart is released when it ends without asking onEnd, so onEnd cannot
   sample it again. The start decision also reaches the span's context. *)
METHOD testOnEndCannotKeepSpanDroppedOnStart : REFERENCE TO FB_Test
VAR
	sampler: FB_Sampler_ForInspection;
	resource: FB_Resource('');
	idGenerator: FB_MockIdGenerator;
	provider: FB_TracerProvider_ForInspection(resource:=resource, idGenerator:=idGenerator, sampler:=sampler);
	scope: FB_InstrumentationScope('sampler.test', '1.0.0', '');
	tracer: FB_Tracer(scope:=scope, provider:=provider);
	processor: FB_SpanProcessor_ForInspection(exporter:=0);
	pSpan: POINTER TO FB_Span;
	pContext: POINTER TO FB_SpanContext;
	ended: BOOL;
END_VAR
TcUnit.TEST('testOnEndCannotKeepSpanDroppedOnStart');
	sampler.dropOnStart := TRUE;
	sampler.sampleOnEnd := TRUE;
	provider.stageProcessor(processor);

	tracer.startSpan(name:='work').build(pDest:=pSpan);
	THIS^.AssertEquals_UDINT(1, sampler.startCount, 'Expected build to call onStart once');
	THIS^.AssertTrue(pSpan <> 0, 'Expected the span to be built');
	IF pSpan <> 0 THEN
		tracer.getSpanContext(pSpan:=pSpan, pDest:=pContext);
		THIS^.AssertTrue(pContext <> 0 AND_THEN (pContext^.traceFlags AND 16#01) = 0, 'Expected the context to carry the start decision');
	END_IF

	ended := tracer.endSpan(pSpan:=pSpan);
	THIS^.AssertTrue(ended, 'Expected endSpan to succeed for a span that is sampled out');
	THIS^.AssertEquals_UDINT(0, sampler.endCount, 'Expected onEnd not to be asked about an unsampled span');
	THIS^.AssertEquals_UDINT(0, provider.spans.count, 'Expected the unsampled span not to be queued');

	provider.tick();
	THIS^.AssertEquals_UDINT(0, processor.exportedCount, 'Expected the unsampled span not to reach the processor');

	IF pContext <> 0 THEN pContext^.delete(pSelf:=pContext); END_IF
TcUnit.TEST_FINISHED();
END_METHOD

(* A root span that only links to an unsampled context is still sampled: a link carries no
   sampling decision into the PLC's trace. *)
METHOD testLinkDoesNotAffectSampling : REFERENCE TO FB_Test
VAR
	resource: FB_Resource('');
	idGenerator: FB_MockIdGenerator;
	provider: FB_TracerProvider_ForInspection(resource:=resource, idGenerator:=idGenerator, sampler:=TcOtlp_GVL.defaultSampler);
	scope: FB_InstrumentationScope('sampler.test', '1.0.0', '');
	tracer: FB_Tracer(scope:=scope, provider:=provider);
	processor: FB_SpanProcessor_ForInspection(exporter:=0);
	unsampled: STRING(55) := '00-4bf92f3577b34da6a3ce929d0e0e4736-00f067aa0ba902b7-00';
	pTrigger: POINTER TO FB_SpanContext;
	pSpan: POINTER TO FB_Span;
END_VAR
TcUnit.TEST('testLinkDoesNotAffectSampling');
	TraceContextPropagator.extract(pDest:=pTrigger, traceparent:=unsampled, tracestate:='');
	THIS^.AssertTrue(pTrigger <> 0, 'Expected the trigger context to be extracted');

	provider.stageProcessor(processor);
	tracer.startSpan(name:='linked.root').addLink(pContext:=pTrigger).build(pDest:=pSpan);
	tracer.endSpan(pSpan:=pSpan);
	provider.tick();

	THIS^.AssertEquals_UDINT(1, processor.exportedCount, 'Expected the linked root span to be processed');

	IF pTrigger <> 0 THEN pTrigger^.delete(pSelf:=pTrigger); END_IF
TcUnit.TEST_FINISHED();
END_METHOD

END_FUNCTION_BLOCK

// ---- TEST/TRACING/SAMPLING/FB_Sampler_ForInspection.TcPOU
(* Sampler test double that counts its calls and can be told to drop spans on start and to
   try to sample them again on end. *)
FUNCTION_BLOCK FB_Sampler_ForInspection EXTENDS FB_Sampler
VAR_INPUT
	dropOnStart: BOOL;  // clear the sampled bit in onStart
	sampleOnEnd: BOOL;  // set the sampled bit in onEnd
END_VAR
VAR_OUTPUT
	startCount: UDINT;
	endCount: UDINT;
END_VAR

METHOD onStart
VAR_INPUT
	span: REFERENCE TO FB_Span;
END_VAR
THIS^.startCount := THIS^.startCount + 1;
SUPER^.onStart(span:=span);
IF THIS^.dropOnStart THEN
	span.setSampled(FALSE);
END_IF
END_METHOD

METHOD onEnd
VAR_INPUT
	span: REFERENCE TO FB_Span;
END_VAR
THIS^.endCount := THIS^.endCount + 1;
IF THIS^.sampleOnEnd THEN
	span.setSampled(TRUE);
END_IF
END_METHOD

END_FUNCTION_BLOCK

// ---- TEST/TRACING/SERIALIZATION/FB_TestSpanProtoJsonSerializer.TcPOU
(* Tests FB_SpanProtoJsonSerializer: span fields, and grouping by resource and scope. *)
FUNCTION_BLOCK FB_TestSpanProtoJsonSerializer EXTENDS FB_TestSuite

THIS^.testSerializeRootSpan();
THIS^.testSerializeChildSpan();
THIS^.testSerializeSpanRejectsInvalidInput();
THIS^.testSerializeTracesDataWithEmptyQueue();
THIS^.testSerializeTracesDataGroupsByResourceAndScope();
THIS^.testSerializeSpanLinks();
THIS^.testSerializeLongTraceState();

(* A root span is written with hex identifiers, numeric enums, string timestamps, attributes and status, and no parentSpanId. *)
METHOD testSerializeRootSpan : REFERENCE TO FB_Test
VAR
	resource: FB_Resource('');
	idGenerator: FB_MockIdGenerator;
	provider: FB_TracerProvider_ForInspection(resource:=resource, idGenerator:=idGenerator, sampler:=TcOtlp_GVL.defaultSampler);
	scope: FB_InstrumentationScope('tracer.test', '1.0.0', '');
	tracer: FB_Tracer(scope:=scope, provider:=provider);
	serializer: FB_SpanProtoJsonSerializer;
	pSpan: POINTER TO FB_Span;
	root: SJsonValue;
	spans: SJsonValue;
	obj: SJsonValue;
	attribute: SJsonValue;
	status: SJsonValue;
	success: BOOL;
	reason: E_ProtoJsonSerializerFailureReason;
END_VAR
TcUnit.TEST('testSerializeRootSpan');
	tracer
		.startSpan(name:='work')
		.setStringAttribute(key:='stats.label', value:='pVal')
		.build(pDest:=pSpan);
	THIS^.AssertTrue(pSpan <> 0, 'Expected the span to build');
	IF pSpan <> 0 THEN
		// no builder sets timestamps; fixed values replace the clock so the output is known
		pSpan^.startTimestamp := 1000;
		pSpan^.endTimestamp := 1581452773000000789;
		tracer.setSpanStatusError(pSpan:=pSpan, message:='motor stalled');

		root := serializer.parser.NewDocument();
		root := serializer.parser.SetObject(root);
		spans := serializer.parser.AddArrayMember(root, 'spans', 0);
		success := serializer.serializeSpan(v:=spans, pSpan:=pSpan, failureReason=>reason);
		THIS^.AssertTrue(success, 'Expected the span to serialize');
		THIS^.AssertEquals_UDINT(TO_UDINT(E_ProtoJsonSerializerFailureReason.NA), TO_UDINT(reason), 'Expected no failure reason');

		obj := serializer.parser.GetArrayValueByIdx(spans, 0);
		THIS^.AssertTrue(serializer.parser.IsObject(obj), 'Expected one Span object');
		// FB_MockIdGenerator fills each new id with one counter byte: the trace id gets 01, the span id 02
		THIS^.AssertEquals_STRING('01010101010101010101010101010101', serializer.parser.GetString(serializer.parser.FindMember(obj, 'traceId')), 'Expected the hex traceId');
		THIS^.AssertEquals_STRING('0202020202020202', serializer.parser.GetString(serializer.parser.FindMember(obj, 'spanId')), 'Expected the hex spanId');
		THIS^.AssertTrue(serializer.parser.FindMember(obj, 'parentSpanId') = 0, 'Expected a root span to omit parentSpanId');
		THIS^.AssertEquals_STRING('work', serializer.parser.GetString(serializer.parser.FindMember(obj, 'name')), 'Expected the name');
		THIS^.AssertEquals_UDINT(1, serializer.parser.GetUint(serializer.parser.FindMember(obj, 'kind')), 'Expected SPAN_KIND_INTERNAL as a number');
		THIS^.AssertEquals_STRING('1000', serializer.parser.GetString(serializer.parser.FindMember(obj, 'startTimeUnixNano')), 'Expected a string startTimeUnixNano');
		THIS^.AssertEquals_STRING('1581452773000000789', serializer.parser.GetString(serializer.parser.FindMember(obj, 'endTimeUnixNano')), 'Expected a string endTimeUnixNano');

		attribute := serializer.parser.GetArrayValueByIdx(serializer.parser.FindMember(obj, 'attributes'), 0);
		THIS^.AssertEquals_STRING('stats.label', serializer.parser.GetString(serializer.parser.FindMember(attribute, 'key')), 'Expected the attribute key');
		THIS^.AssertEquals_STRING(
			'pVal',
			serializer.parser.GetString(serializer.parser.FindMember(serializer.parser.FindMember(attribute, 'value'), 'stringValue')),
			'Expected the attribute value'
		);

		status := serializer.parser.FindMember(obj, 'status');
		THIS^.AssertEquals_UDINT(2, serializer.parser.GetUint(serializer.parser.FindMember(status, 'code')), 'Expected STATUS_CODE_ERROR as a number');
		THIS^.AssertEquals_STRING('motor stalled', serializer.parser.GetString(serializer.parser.FindMember(status, 'message')), 'Expected the status message');
		THIS^.AssertTrue(pSpan^.name <> 0 AND_THEN pSpan^.status <> 0, 'Expected serialization to leave the span intact');
	END_IF

	IF pSpan <> 0 THEN pSpan^.delete(pSelf:=pSpan); END_IF
TcUnit.TEST_FINISHED();
END_METHOD

(* A child span is written with its parentSpanId and kind, and without a status when none is set. *)
METHOD testSerializeChildSpan : REFERENCE TO FB_Test
VAR
	resource: FB_Resource('');
	idGenerator: FB_MockIdGenerator;
	provider: FB_TracerProvider_ForInspection(resource:=resource, idGenerator:=idGenerator, sampler:=TcOtlp_GVL.defaultSampler);
	scope: FB_InstrumentationScope('tracer.test', '1.0.0', '');
	tracer: FB_Tracer(scope:=scope, provider:=provider);
	serializer: FB_SpanProtoJsonSerializer;
	pRoot: POINTER TO FB_Span;
	pChild: POINTER TO FB_Span;
	pContext: POINTER TO FB_SpanContext;
	root: SJsonValue;
	spans: SJsonValue;
	obj: SJsonValue;
	success: BOOL;
END_VAR
TcUnit.TEST('testSerializeChildSpan');
	tracer.startSpan(name:='root').build(pDest:=pRoot);
	IF pRoot <> 0 THEN
		tracer.getSpanContext(pSpan:=pRoot, pDest:=pContext);
	END_IF
	tracer
		.startSpan(name:='child', kind:=E_SpanKind.SPAN_KIND_CLIENT)
		.setParentUsingContext(pContext:=pContext)
		.build(pDest:=pChild);
	THIS^.AssertTrue(pChild <> 0, 'Expected the child span to build');
	IF pChild <> 0 THEN
		root := serializer.parser.NewDocument();
		root := serializer.parser.SetObject(root);
		spans := serializer.parser.AddArrayMember(root, 'spans', 0);
		success := serializer.serializeSpan(v:=spans, pSpan:=pChild);
		THIS^.AssertTrue(success, 'Expected the child span to serialize');

		obj := serializer.parser.GetArrayValueByIdx(spans, 0);
		// FB_MockIdGenerator fills each new id with one counter byte: the root takes trace 01 and
		// span 02, and the child keeps the root's trace and takes span 03
		THIS^.AssertEquals_STRING('0303030303030303', serializer.parser.GetString(serializer.parser.FindMember(obj, 'spanId')), 'Expected the child spanId');
		THIS^.AssertEquals_STRING('0202020202020202', serializer.parser.GetString(serializer.parser.FindMember(obj, 'parentSpanId')), 'Expected the parent spanId');
		THIS^.AssertEquals_UDINT(3, serializer.parser.GetUint(serializer.parser.FindMember(obj, 'kind')), 'Expected SPAN_KIND_CLIENT as a number');
		THIS^.AssertTrue(serializer.parser.FindMember(obj, 'status') = 0, 'Expected no status member');
		THIS^.AssertTrue(serializer.parser.FindMember(obj, 'attributes') = 0, 'Expected no attributes member');
	END_IF

	IF pContext <> 0 THEN pContext^.delete(pSelf:=pContext); END_IF
	IF pChild <> 0 THEN pChild^.delete(pSelf:=pChild); END_IF
	IF pRoot <> 0 THEN pRoot^.delete(pSelf:=pRoot); END_IF
TcUnit.TEST_FINISHED();
END_METHOD

(* serializeSpan reports a null span and an invalid JSON destination. *)
METHOD testSerializeSpanRejectsInvalidInput : REFERENCE TO FB_Test
VAR
	resource: FB_Resource('');
	idGenerator: FB_MockIdGenerator;
	provider: FB_TracerProvider_ForInspection(resource:=resource, idGenerator:=idGenerator, sampler:=TcOtlp_GVL.defaultSampler);
	scope: FB_InstrumentationScope('tracer.test', '1.0.0', '');
	tracer: FB_Tracer(scope:=scope, provider:=provider);
	serializer: FB_SpanProtoJsonSerializer;
	root: SJsonValue;
	spans: SJsonValue;
	invalid: SJsonValue;
	pSpan: POINTER TO FB_Span;
	success: BOOL;
	reason: E_ProtoJsonSerializerFailureReason;
END_VAR
TcUnit.TEST('testSerializeSpanRejectsInvalidInput');
	root := serializer.parser.NewDocument();
	root := serializer.parser.SetObject(root);
	spans := serializer.parser.AddArrayMember(root, 'spans', 0);

	success := serializer.serializeSpan(v:=spans, pSpan:=pSpan, failureReason=>reason);
	THIS^.AssertFalse(success, 'Expected a null span to fail');
	THIS^.AssertEquals_UDINT(TO_UDINT(E_ProtoJsonSerializerFailureReason.SPAN_POINTER_NULL), TO_UDINT(reason), 'Expected SPAN_POINTER_NULL');

	// a valid span, so the only fault left is the destination, which invalid leaves at 0
	tracer.startSpan(name:='work').build(pDest:=pSpan);
	THIS^.AssertTrue(pSpan <> 0, 'Expected the span to build');
	success := serializer.serializeSpan(v:=invalid, pSpan:=pSpan, failureReason=>reason);
	THIS^.AssertFalse(success, 'Expected an invalid destination to fail');
	THIS^.AssertEquals_UDINT(TO_UDINT(E_ProtoJsonSerializerFailureReason.JSON_VALUE_INVALID), TO_UDINT(reason), 'Expected JSON_VALUE_INVALID');
	IF pSpan <> 0 THEN pSpan^.delete(pSelf:=pSpan); END_IF
TcUnit.TEST_FINISHED();
END_METHOD

(* An empty queue gives a document with an empty resourceSpans array. *)
METHOD testSerializeTracesDataWithEmptyQueue : REFERENCE TO FB_Test
VAR
	serializer: FB_SpanProtoJsonSerializer;
	queue: FB_SpanQueue(maxCount:=0);
	resourceSpans: SJsonValue;
	success: BOOL;
	reason: E_ProtoJsonSerializerFailureReason;
END_VAR
TcUnit.TEST('testSerializeTracesDataWithEmptyQueue');
	success := serializer.serializeTracesData(spans:=queue, failureReason=>reason);
	THIS^.AssertTrue(success, 'Expected an empty queue to serialize');
	THIS^.AssertEquals_UDINT(TO_UDINT(E_ProtoJsonSerializerFailureReason.NA), TO_UDINT(reason), 'Expected no failure reason');
	resourceSpans := serializer.parser.FindMember(serializer.jsonValue, 'resourceSpans');
	THIS^.AssertTrue(resourceSpans <> 0 AND_THEN serializer.parser.IsArray(resourceSpans), 'Expected a resourceSpans array');
	THIS^.AssertTrue(serializer.parser.GetArrayValueByIdx(resourceSpans, 0) = 0, 'Expected no ResourceSpans groups');
TcUnit.TEST_FINISHED();
END_METHOD

(*
	Spans arrive with interleaved resources and scopes. Each resource is written once with
	its scopes in first-seen order, and spans keep queue order inside a scope. The serializer
	drains the queue, releasing every span.
*)
METHOD testSerializeTracesDataGroupsByResourceAndScope : REFERENCE TO FB_Test
VAR
	idGenerator: FB_MockIdGenerator;
	resourceB: FB_Resource('resource.b');
	resourceA: FB_Resource('resource.a');
	resourceC: FB_Resource('resource.c');
	providerB: FB_TracerProvider_ForInspection(resource:=resourceB, idGenerator:=idGenerator, sampler:=TcOtlp_GVL.defaultSampler);
	providerA: FB_TracerProvider_ForInspection(resource:=resourceA, idGenerator:=idGenerator, sampler:=TcOtlp_GVL.defaultSampler);
	providerC: FB_TracerProvider_ForInspection(resource:=resourceC, idGenerator:=idGenerator, sampler:=TcOtlp_GVL.defaultSampler);
	scopeB: FB_InstrumentationScope('scope.b', '1.0.0', 'scope.b.schema');
	scopeA: FB_InstrumentationScope('scope.a', '1.0.0', 'scope.a.schema');
	scopeC: FB_InstrumentationScope('scope.c', '1.0.0', 'scope.c.schema');
	tracerBb: FB_Tracer(scope:=scopeB, provider:=providerB);
	tracerBa: FB_Tracer(scope:=scopeA, provider:=providerB);
	tracerAc: FB_Tracer(scope:=scopeC, provider:=providerA);
	tracerAb: FB_Tracer(scope:=scopeB, provider:=providerA);
	tracerCa: FB_Tracer(scope:=scopeA, provider:=providerC);
	queue: FB_SpanQueue(maxCount:=0);
	serializer: FB_SpanProtoJsonSerializer;
	pSpan: POINTER TO FB_Span;
	name: T_MaxString;
	idx: UDINT;
	success: BOOL;
	reason: E_ProtoJsonSerializerFailureReason;
	resourceSpans: SJsonValue;
	resourceObj: SJsonValue;
	scopeSpans: SJsonValue;
	scopeObj: SJsonValue;
	spanArray: SJsonValue;
	spanObj: SJsonValue;
END_VAR
TcUnit.TEST('testSerializeTracesDataGroupsByResourceAndScope');
	// ---- Arrange: eight spans with interleaved resource/scope pairs ----
	// Each tracer is one resource/scope pair, named resource then scope (tracerBa is resource B, scope A).
	// The name holds the span number, so each span can be identified in the output.
	//   span:     1  2  3  4  5  6  7  8
	//   resource: B  A  C  B  C  A  B  A
	//   scope:    B  C  A  A  A  B  B  C
	FOR idx := 1 TO 8 DO
		name := CONCAT('span', UDINT_TO_STRING(idx));
		CASE idx OF
			1, 7: tracerBb.startSpan(name:=name).build(pDest:=pSpan);
			4: tracerBa.startSpan(name:=name).build(pDest:=pSpan);
			2, 8: tracerAc.startSpan(name:=name).build(pDest:=pSpan);
			6: tracerAb.startSpan(name:=name).build(pDest:=pSpan);
			3, 5: tracerCa.startSpan(name:=name).build(pDest:=pSpan);
		END_CASE
		THIS^.AssertTrue(pSpan <> 0, CONCAT('Expected to build ', name));
		IF pSpan <> 0 AND_THEN NOT queue.push(pValue:=pSpan) THEN
			pSpan^.delete(pSelf:=pSpan);
		END_IF
	END_FOR
	THIS^.AssertEquals_UDINT(8, queue.count, 'Expected eight queued spans');

	// ---- Act ----
	success := serializer.serializeTracesData(spans:=queue, failureReason=>reason);
	THIS^.AssertTrue(success, 'Expected TracesData to serialize');
	THIS^.AssertEquals_UDINT(TO_UDINT(E_ProtoJsonSerializerFailureReason.NA), TO_UDINT(reason), 'Expected no failure reason');
	THIS^.AssertEquals_UDINT(0, queue.count, 'Expected the serializer to drain the queue');
	resourceSpans := serializer.parser.FindMember(serializer.jsonValue, 'resourceSpans');
	THIS^.AssertTrue(resourceSpans <> 0 AND_THEN serializer.parser.IsArray(resourceSpans), 'Expected a resourceSpans array');
	THIS^.AssertTrue(serializer.parser.GetArrayValueByIdx(resourceSpans, 3) = 0, 'Expected exactly three ResourceSpans groups');

	// ---- Assert: resource B was seen first, with scope B (spans 1, 7) before scope A (span 4) ----
	resourceObj := serializer.parser.GetArrayValueByIdx(resourceSpans, 0);
	THIS^.AssertEquals_STRING('resource.b', serializer.parser.GetString(serializer.parser.FindMember(resourceObj, 'schemaUrl')), 'Expected resource.b at 0');
	scopeSpans := serializer.parser.FindMember(resourceObj, 'scopeSpans');
	scopeObj := serializer.parser.GetArrayValueByIdx(scopeSpans, 0);
	THIS^.AssertEquals_STRING('scope.b', serializer.parser.GetString(serializer.parser.FindMember(serializer.parser.FindMember(scopeObj, 'scope'), 'name')), 'Expected resource.b scope.b at 0');
	spanArray := serializer.parser.FindMember(scopeObj, 'spans');
	spanObj := serializer.parser.GetArrayValueByIdx(spanArray, 0);
	THIS^.AssertEquals_STRING('span1', serializer.parser.GetString(serializer.parser.FindMember(spanObj, 'name')), 'Expected span1 in resource.b scope.b');
	spanObj := serializer.parser.GetArrayValueByIdx(spanArray, 1);
	THIS^.AssertEquals_STRING('span7', serializer.parser.GetString(serializer.parser.FindMember(spanObj, 'name')), 'Expected span7 in resource.b scope.b');
	THIS^.AssertTrue(serializer.parser.GetArrayValueByIdx(spanArray, 2) = 0, 'Expected 2 span(s) in resource.b scope.b');

	scopeObj := serializer.parser.GetArrayValueByIdx(scopeSpans, 1);
	THIS^.AssertEquals_STRING('scope.a', serializer.parser.GetString(serializer.parser.FindMember(serializer.parser.FindMember(scopeObj, 'scope'), 'name')), 'Expected resource.b scope.a at 1');
	spanArray := serializer.parser.FindMember(scopeObj, 'spans');
	spanObj := serializer.parser.GetArrayValueByIdx(spanArray, 0);
	THIS^.AssertEquals_STRING('span4', serializer.parser.GetString(serializer.parser.FindMember(spanObj, 'name')), 'Expected span4 in resource.b scope.a');
	THIS^.AssertTrue(serializer.parser.GetArrayValueByIdx(spanArray, 1) = 0, 'Expected 1 span(s) in resource.b scope.a');
	THIS^.AssertTrue(serializer.parser.GetArrayValueByIdx(scopeSpans, 2) = 0, 'Expected 2 scope(s) in resource.b');

	// resource A was seen second, with scope C (spans 2, 8) before scope B (span 6)
	resourceObj := serializer.parser.GetArrayValueByIdx(resourceSpans, 1);
	THIS^.AssertEquals_STRING('resource.a', serializer.parser.GetString(serializer.parser.FindMember(resourceObj, 'schemaUrl')), 'Expected resource.a at 1');
	scopeSpans := serializer.parser.FindMember(resourceObj, 'scopeSpans');
	scopeObj := serializer.parser.GetArrayValueByIdx(scopeSpans, 0);
	THIS^.AssertEquals_STRING('scope.c', serializer.parser.GetString(serializer.parser.FindMember(serializer.parser.FindMember(scopeObj, 'scope'), 'name')), 'Expected resource.a scope.c at 0');
	spanArray := serializer.parser.FindMember(scopeObj, 'spans');
	spanObj := serializer.parser.GetArrayValueByIdx(spanArray, 0);
	THIS^.AssertEquals_STRING('span2', serializer.parser.GetString(serializer.parser.FindMember(spanObj, 'name')), 'Expected span2 in resource.a scope.c');
	spanObj := serializer.parser.GetArrayValueByIdx(spanArray, 1);
	THIS^.AssertEquals_STRING('span8', serializer.parser.GetString(serializer.parser.FindMember(spanObj, 'name')), 'Expected span8 in resource.a scope.c');
	THIS^.AssertTrue(serializer.parser.GetArrayValueByIdx(spanArray, 2) = 0, 'Expected 2 span(s) in resource.a scope.c');

	scopeObj := serializer.parser.GetArrayValueByIdx(scopeSpans, 1);
	THIS^.AssertEquals_STRING('scope.b', serializer.parser.GetString(serializer.parser.FindMember(serializer.parser.FindMember(scopeObj, 'scope'), 'name')), 'Expected resource.a scope.b at 1');
	spanArray := serializer.parser.FindMember(scopeObj, 'spans');
	spanObj := serializer.parser.GetArrayValueByIdx(spanArray, 0);
	THIS^.AssertEquals_STRING('span6', serializer.parser.GetString(serializer.parser.FindMember(spanObj, 'name')), 'Expected span6 in resource.a scope.b');
	THIS^.AssertTrue(serializer.parser.GetArrayValueByIdx(spanArray, 1) = 0, 'Expected 1 span(s) in resource.a scope.b');
	THIS^.AssertTrue(serializer.parser.GetArrayValueByIdx(scopeSpans, 2) = 0, 'Expected 2 scope(s) in resource.a');

	// resource C was seen third; its non-adjacent spans 3 and 5 share scope A
	resourceObj := serializer.parser.GetArrayValueByIdx(resourceSpans, 2);
	THIS^.AssertEquals_STRING('resource.c', serializer.parser.GetString(serializer.parser.FindMember(resourceObj, 'schemaUrl')), 'Expected resource.c at 2');
	scopeSpans := serializer.parser.FindMember(resourceObj, 'scopeSpans');
	scopeObj := serializer.parser.GetArrayValueByIdx(scopeSpans, 0);
	THIS^.AssertEquals_STRING('scope.a', serializer.parser.GetString(serializer.parser.FindMember(serializer.parser.FindMember(scopeObj, 'scope'), 'name')), 'Expected resource.c scope.a at 0');
	spanArray := serializer.parser.FindMember(scopeObj, 'spans');
	spanObj := serializer.parser.GetArrayValueByIdx(spanArray, 0);
	THIS^.AssertEquals_STRING('span3', serializer.parser.GetString(serializer.parser.FindMember(spanObj, 'name')), 'Expected span3 in resource.c scope.a');
	spanObj := serializer.parser.GetArrayValueByIdx(spanArray, 1);
	THIS^.AssertEquals_STRING('span5', serializer.parser.GetString(serializer.parser.FindMember(spanObj, 'name')), 'Expected span5 in resource.c scope.a');
	THIS^.AssertTrue(serializer.parser.GetArrayValueByIdx(spanArray, 2) = 0, 'Expected 2 span(s) in resource.c scope.a');
	THIS^.AssertTrue(serializer.parser.GetArrayValueByIdx(scopeSpans, 1) = 0, 'Expected 1 scope(s) in resource.c');

	queue.free();
TcUnit.TEST_FINISHED();
END_METHOD

(* Links are written as a 'links' array in the order they were added, each with hex
   identifiers, flags and any attributes. A span without links writes no 'links' member. *)
METHOD testSerializeSpanLinks : REFERENCE TO FB_Test
VAR
	resource: FB_Resource('');
	idGenerator: FB_MockIdGenerator;
	provider: FB_TracerProvider_ForInspection(resource:=resource, idGenerator:=idGenerator, sampler:=TcOtlp_GVL.defaultSampler);
	scope: FB_InstrumentationScope('tracer.test', '1.0.0', '');
	tracer: FB_Tracer(scope:=scope, provider:=provider);
	serializer: FB_SpanProtoJsonSerializer;
	pTrigger: POINTER TO FB_Span;
	pSpan: POINTER TO FB_Span;
	pTriggerContext: POINTER TO FB_SpanContext;
	pLink: POINTER TO FB_Link;
	root: SJsonValue;
	spans: SJsonValue;
	obj: SJsonValue;
	links: SJsonValue;
	link: SJsonValue;
	attribute: SJsonValue;
	success: BOOL;
	reason: E_ProtoJsonSerializerFailureReason;
END_VAR
TcUnit.TEST('testSerializeSpanLinks');
	tracer.startSpan(name:='trigger').build(pDest:=pTrigger);
	IF pTrigger <> 0 THEN tracer.getSpanContext(pSpan:=pTrigger, pDest:=pTriggerContext); END_IF
	tracer.startSpan(name:='work').addLink(pContext:=pTriggerContext).build(pDest:=pSpan);
	THIS^.AssertTrue(pSpan <> 0, 'Expected the linked span to build');

	// a link with attributes is built with LinkFactory and pushed to the running span
	LinkFactory.fromSpan(pDest:=pLink, pSpan:=pTrigger);
	IF pLink <> 0 THEN
		pLink^.attributes.setStringAttribute(key:='link.reason', value:='retry');
	END_IF
	tracer.pushSpanLink(pSpan:=pSpan, pLink:=pLink);

	IF pSpan <> 0 AND pTrigger <> 0 THEN
		root := serializer.parser.NewDocument();
		root := serializer.parser.SetObject(root);
		spans := serializer.parser.AddArrayMember(root, 'spans', 0);
		success := serializer.serializeSpan(v:=spans, pSpan:=pSpan, failureReason=>reason);
		THIS^.AssertTrue(success, 'Expected the linked span to serialize');
		THIS^.AssertEquals_UDINT(TO_UDINT(E_ProtoJsonSerializerFailureReason.NA), TO_UDINT(reason), 'Expected no failure reason');
		success := serializer.serializeSpan(v:=spans, pSpan:=pTrigger, failureReason=>reason);
		THIS^.AssertTrue(success, 'Expected the trigger span to serialize');

		obj := serializer.parser.GetArrayValueByIdx(spans, 0);
		links := serializer.parser.FindMember(obj, 'links');
		THIS^.AssertTrue(serializer.parser.IsArray(links), 'Expected a links array');
		THIS^.AssertTrue(serializer.parser.FindMember(obj, 'droppedLinksCount') = 0, 'Expected no droppedLinksCount when nothing was dropped');

		link := serializer.parser.GetArrayValueByIdx(links, 0);
		THIS^.AssertTrue(serializer.parser.IsObject(link), 'Expected the first Link object');
		// FB_MockIdGenerator fills each new id with one counter byte: the trigger took trace 01 and span 02
		THIS^.AssertEquals_STRING('01010101010101010101010101010101', serializer.parser.GetString(serializer.parser.FindMember(link, 'traceId')), 'Expected the hex linked traceId');
		THIS^.AssertEquals_STRING('0202020202020202', serializer.parser.GetString(serializer.parser.FindMember(link, 'spanId')), 'Expected the hex linked spanId');
		THIS^.AssertEquals_UDINT(16#101, serializer.parser.GetUint(serializer.parser.FindMember(link, 'flags')), 'Expected the sampled bit and a known local context (16#101)');
		THIS^.AssertTrue(serializer.parser.FindMember(link, 'attributes') = 0, 'Expected no attributes on the first link');
		THIS^.AssertTrue(serializer.parser.FindMember(link, 'traceState') = 0, 'Expected no traceState on the first link');

		link := serializer.parser.GetArrayValueByIdx(links, 1);
		THIS^.AssertTrue(serializer.parser.IsObject(link), 'Expected the second Link object');
		attribute := serializer.parser.GetArrayValueByIdx(serializer.parser.FindMember(link, 'attributes'), 0);
		THIS^.AssertEquals_STRING('link.reason', serializer.parser.GetString(serializer.parser.FindMember(attribute, 'key')), 'Expected the link attribute key');
		THIS^.AssertEquals_STRING(
			'retry',
			serializer.parser.GetString(serializer.parser.FindMember(serializer.parser.FindMember(attribute, 'value'), 'stringValue')),
			'Expected the link attribute value'
		);

		obj := serializer.parser.GetArrayValueByIdx(spans, 1);
		THIS^.AssertTrue(serializer.parser.FindMember(obj, 'links') = 0, 'Expected a span without links to omit links');
	END_IF

	IF pLink <> 0 THEN pLink^.delete(pSelf:=pLink); END_IF
	IF pTriggerContext <> 0 THEN pTriggerContext^.delete(pSelf:=pTriggerContext); END_IF
	IF pSpan <> 0 THEN pSpan^.delete(pSelf:=pSpan); END_IF
	IF pTrigger <> 0 THEN pTrigger^.delete(pSelf:=pTrigger); END_IF
TcUnit.TEST_FINISHED();
END_METHOD

(* A trace state longer than T_MaxString is written whole. W3C asks for at least 512 characters. *)
METHOD testSerializeLongTraceState : REFERENCE TO FB_Test
VAR
	resource: FB_Resource('');
	idGenerator: FB_MockIdGenerator;
	provider: FB_TracerProvider_ForInspection(resource:=resource, idGenerator:=idGenerator, sampler:=TcOtlp_GVL.defaultSampler);
	scope: FB_InstrumentationScope('tracer.test', '1.0.0', '');
	tracer: FB_Tracer(scope:=scope, provider:=provider);
	serializer: FB_SpanProtoJsonSerializer;
	header: STRING(600);
	written: STRING(600);
	pWritten: POINTER TO STRING;
	pBytes: POINTER TO BYTE;
	entry: UDINT;
	i: UDINT;
	n: UDINT;
	traceId: FB_TraceId;
	spanId: FB_SpanId;
	pTraceState: POINTER TO FB_TraceState;
	pRemote: POINTER TO FB_SpanContext;
	pSpan: POINTER TO FB_Span;
	root: SJsonValue;
	spans: SJsonValue;
	obj: SJsonValue;
	member: SJsonValue;
	success: BOOL;
	reason: E_ProtoJsonSerializerFailureReason;
END_VAR
TcUnit.TEST('testSerializeLongTraceState');
	// four 128 character entries joined by ',': 515 characters, built byte by byte
	pBytes := ADR(header);
	FOR entry := 0 TO 3 DO
		IF entry > 0 THEN
			pBytes[n] := 16#2C;  // ','
			n := n + 1;
		END_IF
		pBytes[n] := 16#6B;  // 'k'
		pBytes[n + 1] := 16#30 + TO_BYTE(entry);  // '0' to '3'
		pBytes[n + 2] := 16#3D;  // '='
		n := n + 3;
		FOR i := 1 TO 125 DO  // 125 value characters make a 128 character entry
			pBytes[n] := 16#61 + TO_BYTE(i MOD 26);  // 'a' to 'z'
			n := n + 1;
		END_FOR
	END_FOR
	pBytes[n] := 0;

	MEMSET(ADR(traceId.bytes), 16#AA, SIZEOF(traceId.bytes));
	MEMSET(ADR(spanId.bytes), 16#BB, SIZEOF(spanId.bytes));
	TraceStateFactory.parse(pDest:=pTraceState, pHeader:=ADR(header));
	// 16#301: sampled, remoteness known, remote
	ContextFactory.buildContext(pDest:=pRemote, pTraceId:=ADR(traceId), pSpanId:=ADR(spanId), pTraceState:=pTraceState, traceFlags:=16#301);
	IF pTraceState <> 0 THEN pTraceState^.delete(pSelf:=pTraceState); END_IF
	tracer.startSpan(name:='remote.child').setParentUsingContext(pContext:=pRemote).build(pDest:=pSpan);
	IF pRemote <> 0 THEN pRemote^.delete(pSelf:=pRemote); END_IF
	THIS^.AssertTrue(pSpan <> 0, 'Expected the span to build');

	IF pSpan <> 0 THEN
		root := serializer.parser.NewDocument();
		root := serializer.parser.SetObject(root);
		spans := serializer.parser.AddArrayMember(root, 'spans', 0);
		success := serializer.serializeSpan(v:=spans, pSpan:=pSpan, failureReason=>reason);
		THIS^.AssertTrue(success, 'Expected the span to serialize');

		obj := serializer.parser.GetArrayValueByIdx(spans, 0);
		member := serializer.parser.FindMember(obj, 'traceState');
		THIS^.AssertTrue(member <> 0, 'Expected a traceState member');
		IF member <> 0 THEN
			THIS^.AssertEquals_UDINT(516, TO_UDINT(serializer.parser.GetStringLength(member)), 'Expected all 515 characters and the terminator');
			pWritten := ADR(written);  // CopyString takes a STRING reference and a size, so it can fill a longer buffer
			serializer.parser.CopyString(member, pWritten^, SIZEOF(written));
			THIS^.AssertTrue(MEMCMP(ADR(written), ADR(header), 516) = 0, 'Expected the trace state unchanged');
		END_IF
		pSpan^.delete(pSelf:=pSpan);
	END_IF
TcUnit.TEST_FINISHED();
END_METHOD

END_FUNCTION_BLOCK

// ---- TEST/TRACING/LINK/FB_TestLinks.TcPOU
(* Tests LinkFactory and FB_Links: that a link holds copies of the context it points at, that
   the collection owns its links, keeps their order and refuses links beyond its bound.

   Every test releases the contexts and links it builds before returning. *)
FUNCTION_BLOCK FB_TestLinks EXTENDS FB_TestSuite

THIS^.testFromContextCopiesIdentity();
THIS^.testFromContextRejectsInvalidInput();
THIS^.testFromSpanLinksToTheSpan();
THIS^.testPushTakesOwnershipInOrder();
THIS^.testPushRefusesWhenFull();
THIS^.testFromLinkCopiesLink();
THIS^.testFromLinkRejectsInvalidInput();

(* Builds a span context whose identifier bytes are all seed, for a test to link to. *)
METHOD _buildContext
VAR_IN_OUT
	pDest: POINTER TO FB_SpanContext;
END_VAR
VAR_INPUT
	seed: BYTE;
	traceFlags: UDINT;
END_VAR
VAR
	_traceId: FB_TraceId;
	_spanId: FB_SpanId;
END_VAR
MEMSET(ADR(_traceId.bytes), seed, SIZEOF(_traceId.bytes));
MEMSET(ADR(_spanId.bytes), seed, SIZEOF(_spanId.bytes));
ContextFactory.buildContext(
	pDest:=pDest,
	pTraceId:=ADR(_traceId),
	pSpanId:=ADR(_spanId),
	pTraceState:=0,
	traceFlags:=traceFlags
);
END_METHOD

(* A link holds copies of the context's identity and trace state, so it outlives the context.
   Its flags carry the context's trace flags and remoteness. *)
METHOD testFromContextCopiesIdentity : REFERENCE TO FB_Test
VAR
	pContext: POINTER TO FB_SpanContext;
	pLink: POINTER TO FB_Link;
	traceId: FB_TraceId;
	spanId: FB_SpanId;
	traceStateText: T_MaxString := 'vendor=abc';
	pTraceState: POINTER TO FB_TraceState;
	success: BOOL;
	reason: E_LinkFailureReason;
END_VAR
TcUnit.TEST('testFromContextCopiesIdentity');
	MEMSET(ADR(traceId.bytes), 16#AA, SIZEOF(traceId.bytes));
	MEMSET(ADR(spanId.bytes), 16#BB, SIZEOF(spanId.bytes));
	TraceStateFactory.parse(pDest:=pTraceState, pHeader:=ADR(traceStateText));
	ContextFactory.buildContext(
		pDest:=pContext,
		pTraceId:=ADR(traceId),
		pSpanId:=ADR(spanId),
		pTraceState:=pTraceState,
		traceFlags:=16#301  // sampled, remoteness known, remote
	);
	IF pTraceState <> 0 THEN pTraceState^.delete(pSelf:=pTraceState); END_IF

	success := LinkFactory.fromContext(pDest:=pLink, pContext:=pContext, failureReason=>reason);
	THIS^.AssertTrue(success, 'Expected the link to build');
	THIS^.AssertEquals_UDINT(TO_UDINT(E_LinkFailureReason.NA), TO_UDINT(reason), 'Expected no failure reason');

	// the context is borrowed, so it can be released before the link
	IF pContext <> 0 THEN pContext^.delete(pSelf:=pContext); END_IF

	IF pLink <> 0 THEN
		THIS^.AssertTrue(
			pLink^.traceId <> 0 AND_THEN MEMCMP(ADR(pLink^.traceId^.bytes), ADR(traceId.bytes), SIZEOF(traceId.bytes)) = 0,
			'Expected the linked trace id'
		);
		THIS^.AssertTrue(
			pLink^.spanId <> 0 AND_THEN MEMCMP(ADR(pLink^.spanId^.bytes), ADR(spanId.bytes), SIZEOF(spanId.bytes)) = 0,
			'Expected the linked span id'
		);
		THIS^.AssertTrue(pLink^.traceState <> 0, 'Expected the trace state to be copied');
		IF pLink^.traceState <> 0 THEN
			THIS^.AssertEquals_STRING('vendor=abc', pLink^.traceState^.pString^, 'Expected the trace state text');
		END_IF
		THIS^.AssertEquals_UDINT(16#301, pLink^.flags, 'Expected sampled, remoteness known, remote (16#301)');
		THIS^.AssertEquals_UDINT(0, pLink^.attributes.count, 'Expected no attributes');
		pLink^.delete(pSelf:=pLink);
	END_IF
TcUnit.TEST_FINISHED();
END_METHOD

(* fromContext refuses an assigned destination, a null context and an all zero context,
   and allocates nothing when it does. *)
METHOD testFromContextRejectsInvalidInput : REFERENCE TO FB_Test
VAR
	pContext: POINTER TO FB_SpanContext;
	pZero: POINTER TO FB_SpanContext;
	pLink: POINTER TO FB_Link;
	pOther: POINTER TO FB_Link;
	success: BOOL;
	reason: E_LinkFailureReason;
END_VAR
TcUnit.TEST('testFromContextRejectsInvalidInput');
	THIS^._buildContext(pDest:=pContext, seed:=16#11, traceFlags:=16#101);  // sampled, remoteness known, local
	THIS^._buildContext(pDest:=pZero, seed:=0, traceFlags:=0);  // all zero ids: an invalid context

	success := LinkFactory.fromContext(pDest:=pLink, pContext:=0, failureReason=>reason);
	THIS^.AssertFalse(success, 'Expected a null context to be refused');
	THIS^.AssertEquals_UDINT(TO_UDINT(E_LinkFailureReason.CONTEXT_POINTER_NULL), TO_UDINT(reason), 'Expected CONTEXT_POINTER_NULL');
	THIS^.AssertTrue(pLink = 0, 'Expected nothing to be allocated for a null context');

	success := LinkFactory.fromContext(pDest:=pLink, pContext:=pZero, failureReason=>reason);
	THIS^.AssertFalse(success, 'Expected an invalid context to be refused');
	THIS^.AssertEquals_UDINT(TO_UDINT(E_LinkFailureReason.CONTEXT_INVALID), TO_UDINT(reason), 'Expected CONTEXT_INVALID');
	THIS^.AssertTrue(pLink = 0, 'Expected nothing to be allocated for an invalid context');

	LinkFactory.fromContext(pDest:=pLink, pContext:=pContext);
	pOther := pLink;
	success := LinkFactory.fromContext(pDest:=pLink, pContext:=pContext, failureReason=>reason);
	THIS^.AssertFalse(success, 'Expected an assigned destination to be refused');
	THIS^.AssertEquals_UDINT(TO_UDINT(E_LinkFailureReason.DESTINATION_ALREADY_ASSIGNED), TO_UDINT(reason), 'Expected DESTINATION_ALREADY_ASSIGNED');
	THIS^.AssertTrue(pLink = pOther, 'Expected the destination to be left alone');

	IF pLink <> 0 THEN pLink^.delete(pSelf:=pLink); END_IF
	IF pContext <> 0 THEN pContext^.delete(pSelf:=pContext); END_IF
	IF pZero <> 0 THEN pZero^.delete(pSelf:=pZero); END_IF
TcUnit.TEST_FINISHED();
END_METHOD

(* A link built from a span points at that span, and is local: remoteness is known and not
   remote. A null span is refused. *)
METHOD testFromSpanLinksToTheSpan : REFERENCE TO FB_Test
VAR
	resource: FB_Resource('');
	idGenerator: FB_MockIdGenerator;
	provider: FB_TracerProvider(resource:=resource, idGenerator:=idGenerator, sampler:=TcOtlp_GVL.defaultSampler);
	scope: FB_InstrumentationScope('tracer.test', '1.0.0', '');
	tracer: FB_Tracer(scope:=scope, provider:=provider);
	pSpan: POINTER TO FB_Span;
	pLink: POINTER TO FB_Link;
	success: BOOL;
	reason: E_LinkFailureReason;
END_VAR
TcUnit.TEST('testFromSpanLinksToTheSpan');
	tracer.startSpan(name:='trigger').build(pDest:=pSpan);
	THIS^.AssertTrue(pSpan <> 0, 'Expected the span to build');

	success := LinkFactory.fromSpan(pDest:=pLink, pSpan:=0, failureReason=>reason);
	THIS^.AssertFalse(success, 'Expected a null span to be refused');
	THIS^.AssertEquals_UDINT(TO_UDINT(E_LinkFailureReason.SPAN_POINTER_NULL), TO_UDINT(reason), 'Expected SPAN_POINTER_NULL');

	success := LinkFactory.fromSpan(pDest:=pLink, pSpan:=pSpan, failureReason=>reason);
	THIS^.AssertTrue(success, 'Expected the link to build');
	THIS^.AssertEquals_UDINT(TO_UDINT(E_LinkFailureReason.NA), TO_UDINT(reason), 'Expected no failure reason');
	IF pLink <> 0 AND pSpan <> 0 THEN
		THIS^.AssertTrue(
			MEMCMP(ADR(pLink^.traceId^.bytes), ADR(pSpan^.traceId^.bytes), SIZEOF(pSpan^.traceId^.bytes)) = 0,
			'Expected the span$'s trace id'
		);
		THIS^.AssertTrue(
			MEMCMP(ADR(pLink^.spanId^.bytes), ADR(pSpan^.spanId^.bytes), SIZEOF(pSpan^.spanId^.bytes)) = 0,
			'Expected the span$'s span id'
		);
		THIS^.AssertEquals_UDINT(16#101, pLink^.flags, 'Expected the sampled bit and a known local context (16#101)');
	END_IF

	IF pLink <> 0 THEN pLink^.delete(pSelf:=pLink); END_IF
	IF pSpan <> 0 THEN pSpan^.delete(pSelf:=pSpan); END_IF
TcUnit.TEST_FINISHED();
END_METHOD

(* push takes ownership and clears the caller's pointer; next walks the links oldest first
   without taking them, and pop hands them back in the same order. *)
METHOD testPushTakesOwnershipInOrder : REFERENCE TO FB_Test
VAR
	links: FB_Links(maxCount:=TcOtlp_GVL.DEFAULT_MAX_LINK_COUNT);
	pFirst: POINTER TO FB_SpanContext;
	pSecond: POINTER TO FB_SpanContext;
	pLink: POINTER TO FB_Link;
	pWalked: POINTER TO FB_Link;
	success: BOOL;
	reason: E_LinkFailureReason;
END_VAR
TcUnit.TEST('testPushTakesOwnershipInOrder');
	// 16#101: sampled, remoteness known, local; the seed byte tells the links apart
	THIS^._buildContext(pDest:=pFirst, seed:=16#11, traceFlags:=16#101);
	THIS^._buildContext(pDest:=pSecond, seed:=16#22, traceFlags:=16#101);

	LinkFactory.fromContext(pDest:=pLink, pContext:=pFirst);
	success := links.push(pValue:=pLink, failureReason=>reason);
	THIS^.AssertTrue(success, 'Expected the first push to succeed');
	THIS^.AssertEquals_UDINT(TO_UDINT(E_LinkFailureReason.NA), TO_UDINT(reason), 'Expected no failure reason');
	THIS^.AssertTrue(pLink = 0, 'Expected push to clear the caller$'s pointer');
	LinkFactory.fromContext(pDest:=pLink, pContext:=pSecond);
	links.push(pValue:=pLink);
	THIS^.AssertEquals_UDINT(2, links.count, 'Expected two links');

	links.reset();
	pWalked := links.next();
	THIS^.AssertTrue(pWalked <> 0 AND_THEN pWalked^.spanId^.bytes[0] = 16#11, 'Expected next to start at the oldest link');
	pWalked := links.next();
	THIS^.AssertTrue(pWalked <> 0 AND_THEN pWalked^.spanId^.bytes[0] = 16#22, 'Expected next to reach the second link');
	THIS^.AssertTrue(links.next() = 0, 'Expected next to end after the last link');
	THIS^.AssertEquals_UDINT(2, links.count, 'Expected walking to leave the links in place');

	success := links.pop(pValue:=pLink, failureReason=>reason);
	THIS^.AssertTrue(success AND_THEN pLink^.spanId^.bytes[0] = 16#11, 'Expected pop to return the oldest link');
	success := links.pop(pValue:=pLink, failureReason=>reason);
	THIS^.AssertFalse(success, 'Expected pop into an assigned destination to fail');
	THIS^.AssertEquals_UDINT(TO_UDINT(E_LinkFailureReason.DESTINATION_ALREADY_ASSIGNED), TO_UDINT(reason), 'Expected DESTINATION_ALREADY_ASSIGNED');
	IF pLink <> 0 THEN pLink^.delete(pSelf:=pLink); END_IF

	links.pop(pValue:=pLink);
	IF pLink <> 0 THEN pLink^.delete(pSelf:=pLink); END_IF
	success := links.pop(pValue:=pLink, failureReason=>reason);
	THIS^.AssertFalse(success, 'Expected pop from an empty collection to fail');
	THIS^.AssertEquals_UDINT(TO_UDINT(E_LinkFailureReason.LINKS_EMPTY), TO_UDINT(reason), 'Expected LINKS_EMPTY');
	THIS^.AssertEquals_UDINT(0, links.count, 'Expected no links left');

	IF pFirst <> 0 THEN pFirst^.delete(pSelf:=pFirst); END_IF
	IF pSecond <> 0 THEN pSecond^.delete(pSelf:=pSecond); END_IF
TcUnit.TEST_FINISHED();
END_METHOD

(* A full collection keeps its links and refuses the new one: the caller keeps it, and it is
   counted as dropped. A null link is refused without being counted. free releases every link. *)
METHOD testPushRefusesWhenFull : REFERENCE TO FB_Test
VAR
	links: FB_Links(maxCount:=1);
	pContext: POINTER TO FB_SpanContext;
	pLink: POINTER TO FB_Link;
	pRefused: POINTER TO FB_Link;
	success: BOOL;
	reason: E_LinkFailureReason;
END_VAR
TcUnit.TEST('testPushRefusesWhenFull');
	THIS^._buildContext(pDest:=pContext, seed:=16#11, traceFlags:=16#101);  // sampled, remoteness known, local

	success := links.push(pValue:=pLink, failureReason=>reason);
	THIS^.AssertFalse(success, 'Expected a null link to be refused');
	THIS^.AssertEquals_UDINT(TO_UDINT(E_LinkFailureReason.LINK_POINTER_NULL), TO_UDINT(reason), 'Expected LINK_POINTER_NULL');

	LinkFactory.fromContext(pDest:=pLink, pContext:=pContext);
	links.push(pValue:=pLink);
	LinkFactory.fromContext(pDest:=pLink, pContext:=pContext);
	pRefused := pLink;
	success := links.push(pValue:=pLink, failureReason=>reason);
	THIS^.AssertFalse(success, 'Expected a push beyond maxCount to fail');
	THIS^.AssertEquals_UDINT(TO_UDINT(E_LinkFailureReason.LINK_COUNT_LIMIT_REACHED), TO_UDINT(reason), 'Expected LINK_COUNT_LIMIT_REACHED');
	THIS^.AssertTrue(pLink = pRefused, 'Expected the caller to keep the refused link');
	THIS^.AssertEquals_UDINT(1, links.count, 'Expected the first link to be kept');
	THIS^.AssertEquals_UDINT(1, links.droppedCount, 'Expected the refused link to be counted');
	IF pLink <> 0 THEN pLink^.delete(pSelf:=pLink); END_IF

	THIS^.AssertTrue(links.free(), 'Expected free to release every link');
	THIS^.AssertEquals_UDINT(0, links.count, 'Expected no links after free');
	THIS^.AssertEquals_UDINT(0, links.droppedCount, 'Expected free to clear droppedCount');

	IF pContext <> 0 THEN pContext^.delete(pSelf:=pContext); END_IF
TcUnit.TEST_FINISHED();
END_METHOD

(* fromLink gives the copy its own identity, trace state and attributes. *)
METHOD testFromLinkCopiesLink : REFERENCE TO FB_Test
VAR
	pContext: POINTER TO FB_SpanContext;
	pLink: POINTER TO FB_Link;
	pCopy: POINTER TO FB_Link;
	reason: E_LinkFailureReason;
END_VAR
TcUnit.TEST('testFromLinkCopiesLink');
	THIS^._buildContext(pDest:=pContext, seed:=5, traceFlags:=1);  // sampled only
	LinkFactory.fromContext(pDest:=pLink, pContext:=pContext, failureReason=>reason);
	THIS^.AssertTrue(pLink <> 0, 'Expected the source link to build');
	IF pLink <> 0 THEN
		pLink^.attributes.setStringAttribute('k', 'v');
		THIS^.AssertTrue(LinkFactory.fromLink(pDest:=pCopy, pSrc:=pLink, failureReason=>reason), 'Expected fromLink to succeed');
		IF pCopy <> 0 THEN
			THIS^.AssertTrue(pCopy^.traceId <> 0 AND_THEN pCopy^.traceId <> pLink^.traceId, 'Expected a copied trace id');
			THIS^.AssertTrue(pCopy^.spanId <> 0 AND_THEN pCopy^.spanId <> pLink^.spanId, 'Expected a copied span id');
			THIS^.AssertEquals_UDINT(pLink^.flags, pCopy^.flags, 'Expected the flags');
			THIS^.AssertEquals_UDINT(1, pCopy^.attributes.count, 'Expected the attribute');
			pLink^.delete(pSelf:=pLink);
			THIS^.AssertTrue(pCopy^.traceId^.bytes[0] = 5 AND pCopy^.spanId^.bytes[0] = 5, 'Expected the identity to outlive the source');
			pCopy^.delete(pSelf:=pCopy);
		END_IF
		IF pLink <> 0 THEN pLink^.delete(pSelf:=pLink); END_IF
	END_IF
	IF pContext <> 0 THEN pContext^.delete(pSelf:=pContext); END_IF
TcUnit.TEST_FINISHED();
END_METHOD

(* fromLink refuses a missing source and an assigned destination. *)
METHOD testFromLinkRejectsInvalidInput : REFERENCE TO FB_Test
VAR
	pLink: POINTER TO FB_Link;
	pDest: POINTER TO FB_Link;
	reason: E_LinkFailureReason;
END_VAR
TcUnit.TEST('testFromLinkRejectsInvalidInput');
	THIS^.AssertFalse(LinkFactory.fromLink(pDest:=pDest, pSrc:=0, failureReason=>reason), 'Expected a null source to fail');
	THIS^.AssertEquals_UDINT(TO_UDINT(E_LinkFailureReason.LINK_POINTER_NULL), TO_UDINT(reason), 'Expected LINK_POINTER_NULL');

	pLink := __NEW(FB_Link);  // built by hand: LinkFactory refuses a link with no identity
	THIS^.AssertFalse(LinkFactory.fromLink(pDest:=pDest, pSrc:=pLink, failureReason=>reason), 'Expected an empty link to fail');
	THIS^.AssertEquals_UDINT(TO_UDINT(E_LinkFailureReason.CONTEXT_INVALID), TO_UDINT(reason), 'Expected CONTEXT_INVALID');

	pDest := pLink;
	THIS^.AssertFalse(LinkFactory.fromLink(pDest:=pDest, pSrc:=pLink, failureReason=>reason), 'Expected an assigned destination to fail');
	THIS^.AssertEquals_UDINT(
		TO_UDINT(E_LinkFailureReason.DESTINATION_ALREADY_ASSIGNED),
		TO_UDINT(reason),
		'Expected DESTINATION_ALREADY_ASSIGNED'
	);
	THIS^.AssertTrue(pDest = pLink, 'Expected the destination to be left alone');
	IF pLink <> 0 THEN pLink^.delete(pSelf:=pLink); END_IF
TcUnit.TEST_FINISHED();
END_METHOD

END_FUNCTION_BLOCK

// ---- TEST/TRACING/EXPORTING/FB_TestSpanFileExporter.TcPOU
(*
	Tests FB_SpanExporter_File across scan cycles: it refuses a batch while busy, appends a batch
	to its file, and delivers a second batch handed over right after the first one finished.
*)
FUNCTION_BLOCK FB_TestSpanFileExporter EXTENDS FB_TestSuite
VAR
	_exporter: FB_SpanExporter_File(filepath:='C:\Users\samue\Desktop\programming projects\TcOtlp\spans.jsonl');
	_spans: FB_SpanQueue(maxCount:=0);
	_resource: FB_Resource('');
	_idGenerator: FB_MockIdGenerator;
	_provider: FB_TracerProvider_ForInspection(resource:=_resource, idGenerator:=_idGenerator, sampler:=TcOtlp_GVL.defaultSampler);
	_scope: FB_InstrumentationScope('tracer.test', '1.0.0', '');
	_tracer: FB_Tracer(scope:=_scope, provider:=_provider);
END_VAR

THIS^.testExportWritesSpansToFile();

(*
	The file exporter refuses a second batch while it is busy, leaving the spans with the caller,
	writes an accepted batch to its file, and accepts the next batch in the scan the first one finished.
*)
METHOD testExportWritesSpansToFile : REFERENCE TO FB_Test
VAR CONSTANT
	FILEPATH: STRING := 'C:\Users\samue\Desktop\programming projects\TcOtlp\spans.jsonl';
	MAX_CYCLES: UDINT := 1000;
END_VAR
VAR_INST
	_state: USINT;
	_cycles: UDINT;
	_delivered: UDINT;
	_fileFinder: FB_EnumFindFileEntry;
	_fileDeleter: FB_FileDelete;
END_VAR
VAR
	pSpan: POINTER TO FB_Span;
	idx: UDINT;
	queueReason: E_SpanQueueFailureReason;
	exportReason: E_SpanExporterFailureReason;
	tickSucceeded: BOOL;
END_VAR
TcUnit.TEST('testExportWritesSpansToFile');
	CASE _state OF
		0: // hand over a batch of two spans, then offer another while busy
			_cycles := 0;
			_delivered := 0;
			FOR idx := 1 TO 2 DO
				_tracer.startSpan(name:='work').setStringAttribute(key:='k', value:='v').build(pDest:=pSpan);
				_spans.push(pValue:=pSpan, failureReason=>queueReason);
				IF pSpan <> 0 THEN pSpan^.delete(pSelf:=pSpan); END_IF
			END_FOR
			THIS^.AssertEquals_UDINT(2, _spans.count, 'Expected two queued spans');
			THIS^.AssertTrue(_exporter.export(spans:=_spans, count:=_spans.count, failureReason=>exportReason), 'Expected the exporter to accept the batch');
			THIS^.AssertEquals_UDINT(0, _spans.count, 'Expected the batch to move into the exporter');
			THIS^.AssertTrue(_exporter.isBusy(), 'Expected the exporter to be busy');

			_tracer.startSpan(name:='late').build(pDest:=pSpan);
			_spans.push(pValue:=pSpan, failureReason=>queueReason);
			IF pSpan <> 0 THEN pSpan^.delete(pSelf:=pSpan); END_IF
			THIS^.AssertFalse(_exporter.export(spans:=_spans, count:=1, failureReason=>exportReason), 'Expected a busy exporter to refuse');
			THIS^.AssertEquals_UDINT(
				TO_UDINT(E_SpanExporterFailureReason.ACTIVE_EXPORT_IN_PROGRESS),
				TO_UDINT(exportReason),
				'Expected ACTIVE_EXPORT_IN_PROGRESS'
			);
			THIS^.AssertEquals_UDINT(1, _spans.count, 'Expected the refused span to stay with the caller');
			_spans.free();
			_state := 10;

		10: // deliver the batch, then hand over a second one in the scan it finished
			tickSucceeded := _exporter.tick(failureReason=>exportReason);
			_cycles := _cycles + 1;
			IF NOT tickSucceeded THEN
				THIS^.AssertEquals_UDINT(0, TO_UDINT(exportReason), 'Expected the file export to succeed');
				_state := 30;
			ELSIF _exporter.currentState = E_FileExporterState.done THEN
				THIS^.AssertFalse(_exporter.isBusy(), 'Expected the exporter to release the delivered batch');
				_delivered := _delivered + 1;
				IF _delivered = 1 THEN
					_tracer.startSpan(name:='next').build(pDest:=pSpan);
					_spans.push(pValue:=pSpan, failureReason=>queueReason);
					IF pSpan <> 0 THEN pSpan^.delete(pSelf:=pSpan); END_IF
					THIS^.AssertTrue(_exporter.export(spans:=_spans, count:=1, failureReason=>exportReason), 'Expected a finished exporter to accept the next batch');
					_cycles := 0;
				ELSE
					_state := 20;
				END_IF
			ELSIF _cycles > MAX_CYCLES THEN
				THIS^.AssertTrue(FALSE, 'Expected the file export to finish within MAX_CYCLES');
				_state := 30;
			END_IF

		20: // the batch made the file non-empty
			_fileFinder(sPathName:=FILEPATH, bExecute:=TRUE);
			IF NOT _fileFinder.bBusy THEN
				THIS^.AssertTrue(ULARGE_TO_ULINT(_fileFinder.stFindFile.fileSize) > 0, 'Expected a non-empty file');
				_fileFinder(bExecute:=FALSE);
				_state := 30;
			END_IF

		30: // remove the file
			_fileDeleter(sPathName:=FILEPATH, bExecute:=TRUE);
			IF NOT _fileDeleter.bBusy THEN
				_fileDeleter(bExecute:=FALSE);
				_spans.free();
				_state := 0;
				TcUnit.TEST_FINISHED();
			END_IF
	END_CASE
END_METHOD

END_FUNCTION_BLOCK

// ---- TEST/TRACING/EXPORTING/FB_TestSpanConsoleExporter.TcPOU
(* Tests FB_SpanExporter_Console: the line it writes per span, and that it releases each batch at once. *)
FUNCTION_BLOCK FB_TestSpanConsoleExporter EXTENDS FB_TestSuite

THIS^.testFormatsRootSpan();
THIS^.testFormatsChildSpan();
THIS^.testExportWritesAndReleasesBatch();
THIS^.testSimpleProcessorExportsEverySpan();

(* A root span is written with its identifiers in hex, no parent and its duration. *)
METHOD testFormatsRootSpan : REFERENCE TO FB_Test
VAR
	resource: FB_Resource('');
	idGenerator: FB_MockIdGenerator;
	provider: FB_TracerProvider_ForInspection(resource:=resource, idGenerator:=idGenerator, sampler:=TcOtlp_GVL.defaultSampler);
	scope: FB_InstrumentationScope('tracer.test', '1.0.0', '');
	tracer: FB_Tracer(scope:=scope, provider:=provider);
	exporter: FB_SpanExporter_Console;
	pSpan: POINTER TO FB_Span;
END_VAR
TcUnit.TEST('testFormatsRootSpan');
	tracer.startSpan(name:='work').build(pDest:=pSpan);
	THIS^.AssertTrue(pSpan <> 0, 'Expected the span to build');
	IF pSpan <> 0 THEN
		// the builder has no timestamp setter; fixed values keep the output deterministic
		pSpan^.startTimestamp := 1000;
		pSpan^.endTimestamp := 1500;
		// FB_MockIdGenerator fills each new id with the next counter byte:
		// the trace id is 16#01 repeated, then the span id is 16#02 repeated
		THIS^.AssertEquals_STRING(
			'span "work" trace=01010101010101010101010101010101 span=0202020202020202 parent=none kind=SPAN_KIND_INTERNAL status=STATUS_CODE_UNSET duration=500ns',
			exporter.format(pSpan^),
			'Expected the root span line'
		);
		pSpan^.delete(pSelf:=pSpan);
	END_IF
TcUnit.TEST_FINISHED();
END_METHOD

(* A child span is written with its parent span id and its kind. *)
METHOD testFormatsChildSpan : REFERENCE TO FB_Test
VAR
	resource: FB_Resource('');
	idGenerator: FB_MockIdGenerator;
	provider: FB_TracerProvider_ForInspection(resource:=resource, idGenerator:=idGenerator, sampler:=TcOtlp_GVL.defaultSampler);
	scope: FB_InstrumentationScope('tracer.test', '1.0.0', '');
	tracer: FB_Tracer(scope:=scope, provider:=provider);
	exporter: FB_SpanExporter_Console;
	pRoot: POINTER TO FB_Span;
	pChild: POINTER TO FB_Span;
	pContext: POINTER TO FB_SpanContext;
END_VAR
TcUnit.TEST('testFormatsChildSpan');
	tracer.startSpan(name:='root').build(pDest:=pRoot);
	IF pRoot <> 0 THEN
		tracer.getSpanContext(pSpan:=pRoot, pDest:=pContext);
	END_IF
	tracer
		.startSpan(name:='child', kind:=E_SpanKind.SPAN_KIND_CLIENT)
		.setParentUsingContext(pContext:=pContext)
		.build(pDest:=pChild);
	THIS^.AssertTrue(pChild <> 0, 'Expected the child span to build');
	IF pChild <> 0 THEN
		// the builder has no timestamp setter; fixed values keep the output deterministic
		pChild^.startTimestamp := 2000;
		pChild^.endTimestamp := 2000;
		// FB_MockIdGenerator fills each new id with the next counter byte: the root takes
		// trace id 16#01 and span id 16#02, and the child shares the trace and takes span id 16#03
		THIS^.AssertEquals_STRING(
			'span "child" trace=01010101010101010101010101010101 span=0303030303030303 parent=0202020202020202 kind=SPAN_KIND_CLIENT status=STATUS_CODE_UNSET duration=0ns',
			exporter.format(pChild^),
			'Expected the child span line'
		);
	END_IF

	IF pContext <> 0 THEN pContext^.delete(pSelf:=pContext); END_IF
	IF pChild <> 0 THEN pChild^.delete(pSelf:=pChild); END_IF
	IF pRoot <> 0 THEN pRoot^.delete(pSelf:=pRoot); END_IF
TcUnit.TEST_FINISHED();
END_METHOD

(* export takes the whole batch, writes it and releases it at once, so the exporter is never busy. *)
METHOD testExportWritesAndReleasesBatch : REFERENCE TO FB_Test
VAR
	resource: FB_Resource('');
	idGenerator: FB_MockIdGenerator;
	provider: FB_TracerProvider_ForInspection(resource:=resource, idGenerator:=idGenerator, sampler:=TcOtlp_GVL.defaultSampler);
	scope: FB_InstrumentationScope('tracer.test', '1.0.0', '');
	tracer: FB_Tracer(scope:=scope, provider:=provider);
	exporter: FB_SpanExporter_Console;
	spans: FB_SpanQueue(maxCount:=0);
	pSpan: POINTER TO FB_Span;
	idx: UDINT;
	queueReason: E_SpanQueueFailureReason;
	exportReason: E_SpanExporterFailureReason;
END_VAR
TcUnit.TEST('testExportWritesAndReleasesBatch');
	FOR idx := 1 TO 2 DO
		tracer.startSpan(name:='work').build(pDest:=pSpan);
		spans.push(pValue:=pSpan, failureReason=>queueReason);
		IF pSpan <> 0 THEN pSpan^.delete(pSelf:=pSpan); END_IF
	END_FOR
	THIS^.AssertEquals_UDINT(2, spans.count, 'Expected two queued spans');

	THIS^.AssertTrue(exporter.export(spans:=spans, count:=spans.count, failureReason=>exportReason), 'Expected the exporter to accept the batch');
	THIS^.AssertEquals_UDINT(0, TO_UDINT(exportReason), 'Expected no failure');
	THIS^.AssertEquals_UDINT(0, spans.count, 'Expected the batch to move into the exporter');
	THIS^.AssertFalse(exporter.isBusy(), 'Expected the exporter to release the batch before returning');
	THIS^.AssertTrue(exporter.tick(failureReason=>exportReason), 'Expected tick to succeed');
	spans.free();
TcUnit.TEST_FINISHED();
END_METHOD

(* A simple processor with a console exporter writes every span, even spans ending in the same scan. *)
METHOD testSimpleProcessorExportsEverySpan : REFERENCE TO FB_Test
VAR
	resource: FB_Resource('');
	idGenerator: FB_MockIdGenerator;
	provider: FB_TracerProvider_ForInspection(resource:=resource, idGenerator:=idGenerator, sampler:=TcOtlp_GVL.defaultSampler);
	scope: FB_InstrumentationScope('tracer.test', '1.0.0', '');
	tracer: FB_Tracer(scope:=scope, provider:=provider);
	exporter: FB_SpanExporter_Console;
	processor: FB_SpanProcessor_Simple(exporter:=exporter);
	pSpan: POINTER TO FB_Span;
	idx: UDINT;
END_VAR
TcUnit.TEST('testSimpleProcessorExportsEverySpan');
	FOR idx := 1 TO 2 DO
		tracer.startSpan(name:='work').build(pDest:=pSpan);
		THIS^.AssertTrue(pSpan <> 0, 'Expected the span to build');
		IF pSpan <> 0 THEN
			THIS^.AssertFalse(exporter.isBusy(), 'Expected the console exporter to be free for every span');
			processor.onEnd(pSpan^);  // writes the line to the ADS log
			pSpan^.delete(pSelf:=pSpan);
		END_IF
	END_FOR
	THIS^.AssertFalse(exporter.isBusy(), 'Expected the console exporter to hold no batch');
TcUnit.TEST_FINISHED();
END_METHOD

END_FUNCTION_BLOCK

// ---- TEST/TRACING/EXPORTING/FB_TestSpanHttpExporter.TcPOU
(*
	Tests FB_SpanExporter_HTTP without a collector: an invalid URL fails at once, a refused
	connection is reported as HTTP_REQUEST_FAILURE, and a failed exporter accepts and starts
	the next batch.
*)
FUNCTION_BLOCK FB_TestSpanHttpExporter EXTENDS FB_TestSuite
VAR
	_exporterBadUrl: FB_SpanExporter_HTTP(url:='not-a-valid-url', bNoServerCertCheck:=TRUE);
	_exporterRefused: FB_SpanExporter_HTTP(url:='http://127.0.0.1:1/v1/traces', bNoServerCertCheck:=TRUE);
	_spans: FB_SpanQueue(maxCount:=0);
	_resource: FB_Resource('');
	_idGenerator: FB_MockIdGenerator;
	_provider: FB_TracerProvider_ForInspection(resource:=_resource, idGenerator:=_idGenerator, sampler:=TcOtlp_GVL.defaultSampler);
	_scope: FB_InstrumentationScope('tracer.test', '1.0.0', '');
	_tracer: FB_Tracer(scope:=_scope, provider:=_provider);
END_VAR

THIS^.testInvalidUrlFailsFast();
THIS^.testConnectionRefusedReportsFailure();

(* Builds a span and queues a copy of it in _spans. *)
METHOD queueSpan
VAR_INPUT
	name: STRING;
END_VAR
VAR
	pSpan: POINTER TO FB_Span;
	queueReason: E_SpanQueueFailureReason;
END_VAR
_tracer.startSpan(name:=name).build(pDest:=pSpan);
THIS^._spans.push(pValue:=pSpan, failureReason=>queueReason);
IF pSpan <> 0 THEN pSpan^.delete(pSelf:=pSpan); END_IF
END_METHOD

(* An unparseable URL fails in the first tick without sending, and the batch is released. *)
METHOD testInvalidUrlFailsFast : REFERENCE TO FB_Test
VAR
	exportReason: E_SpanExporterFailureReason;
END_VAR
TcUnit.TEST('testInvalidUrlFailsFast');
	THIS^.queueSpan('work');
	THIS^.AssertEquals_UDINT(1, _spans.count, 'Expected one queued span');
	THIS^.AssertTrue(_exporterBadUrl.export(spans:=_spans, count:=1, failureReason=>exportReason), 'Expected the exporter to accept the batch before checking the URL');
	THIS^.AssertEquals_UDINT(0, _spans.count, 'Expected the batch to move into the exporter');
	THIS^.AssertTrue(_exporterBadUrl.isBusy(), 'Expected the exporter to be busy');

